// TIA Portal V20 program export: 0 tag tables, 36 data types, 10 data blocks, 80 code blocks (in call order from the OBs), 3 instance data blocks

TYPE "FRK_Access"
// stored: IsFailsafeCompliant false
   STRUCT
      CurrentLevel : DInt;
      CurrentUser : String[32];
      LoginFailed : Bool;
      Policy { S7_SetPoint := 'True'} : "ST_AccessPolicy";
      SessionGeneration : UDInt;
      LoginBusy : Bool;
      LoginResultSequence : UDInt;
      LoginTimeoutMs : UDInt;
      ProviderEnabled { ExternalAccessible := 'False'; ExternalVisible := 'False'; ExternalWritable := 'False'} : Bool;
      LastActivity { ExternalAccessible := 'False'; ExternalVisible := 'False'; ExternalWritable := 'False'} : UDInt;
      LoginSince { ExternalAccessible := 'False'; ExternalVisible := 'False'; ExternalWritable := 'False'} : UDInt;
      LoginSequence { ExternalAccessible := 'False'; ExternalVisible := 'False'; ExternalWritable := 'False'} : UDInt;
      CandidateUser { ExternalAccessible := 'False'; ExternalVisible := 'False'; ExternalWritable := 'False'} : String[32];
      CandidateLevel { ExternalAccessible := 'False'; ExternalVisible := 'False'; ExternalWritable := 'False'} : DInt;
      Round { ExternalAccessible := 'False'; ExternalVisible := 'False'; ExternalWritable := 'False'} : DInt;
      Salt { ExternalAccessible := 'False'; ExternalVisible := 'False'; ExternalWritable := 'False'} : Array[0..15] of Byte;
      Digest { ExternalAccessible := 'False'; ExternalVisible := 'False'; ExternalWritable := 'False'} : Array[0..31] of Byte;
      Expected { ExternalAccessible := 'False'; ExternalVisible := 'False'; ExternalWritable := 'False'} : Array[0..31] of Byte;
   END_STRUCT;
END_TYPE

TYPE "FRK_Carrier"
// stored: IsFailsafeCompliant false
   STRUCT
      Enabled { ExternalAccessible := 'False'; ExternalVisible := 'False'; ExternalWritable := 'False'} : Bool;
      Kind { ExternalAccessible := 'False'; ExternalVisible := 'False'; ExternalWritable := 'False'} : DInt;
      Serial { ExternalAccessible := 'False'; ExternalVisible := 'False'; ExternalWritable := 'False'} : UDInt;
      Context { ExternalAccessible := 'False'; ExternalVisible := 'False'; ExternalWritable := 'False'; S7_SetPoint := 'True'} : "ST_PartContext";
      Written { ExternalAccessible := 'False'; ExternalVisible := 'False'; ExternalWritable := 'False'; S7_SetPoint := 'True'} : "ST_PartContext";
      Writes { ExternalAccessible := 'False'; ExternalVisible := 'False'; ExternalWritable := 'False'} : UDInt;
   END_STRUCT;
END_TYPE

TYPE "FRK_ConfigCursor"
// stored: IsFailsafeCompliant false
   STRUCT
      Position { ExternalAccessible := 'False'; ExternalVisible := 'False'; ExternalWritable := 'False'} : DInt;
      First { ExternalAccessible := 'False'; ExternalVisible := 'False'; ExternalWritable := 'False'} : DInt;
   END_STRUCT;
END_TYPE

TYPE "FRK_Core"
// stored: IsFailsafeCompliant false
   STRUCT
      Named { ExternalAccessible := 'False'; ExternalVisible := 'False'; ExternalWritable := 'False'} : Bool;
      Initialized { ExternalAccessible := 'False'; ExternalVisible := 'False'; ExternalWritable := 'False'} : Bool;
      RegIndex { ExternalAccessible := 'False'; ExternalVisible := 'False'; ExternalWritable := 'False'} : DInt;
      ParentIndex { ExternalAccessible := 'False'; ExternalVisible := 'False'; ExternalWritable := 'False'} : DInt;
      ModuleType { ExternalAccessible := 'False'; ExternalVisible := 'False'; ExternalWritable := 'False'} : DInt;
      Exec { ExternalAccessible := 'False'; ExternalVisible := 'False'; ExternalWritable := 'False'} : DInt;
      ExecPrev { ExternalAccessible := 'False'; ExternalVisible := 'False'; ExternalWritable := 'False'} : Bool;
      AbortPrev { ExternalAccessible := 'False'; ExternalVisible := 'False'; ExternalWritable := 'False'} : Bool;
      Armed { ExternalAccessible := 'False'; ExternalVisible := 'False'; ExternalWritable := 'False'} : Bool;
      Command { ExternalAccessible := 'False'; ExternalVisible := 'False'; ExternalWritable := 'False'} : DInt;
      CommandLabel { ExternalAccessible := 'False'; ExternalVisible := 'False'; ExternalWritable := 'False'} : String[120];
      Dispatch { ExternalAccessible := 'False'; ExternalVisible := 'False'; ExternalWritable := 'False'} : Bool;
      EvInit { ExternalAccessible := 'False'; ExternalVisible := 'False'; ExternalWritable := 'False'} : Bool;
      EvCommandStart { ExternalAccessible := 'False'; ExternalVisible := 'False'; ExternalWritable := 'False'} : Bool;
      ReleasePending { ExternalAccessible := 'False'; ExternalVisible := 'False'; ExternalWritable := 'False'} : Bool;
      EvAbort { ExternalAccessible := 'False'; ExternalVisible := 'False'; ExternalWritable := 'False'} : Bool;
      EvAbortInError { ExternalAccessible := 'False'; ExternalVisible := 'False'; ExternalWritable := 'False'} : Bool;
      EvModeExit { ExternalAccessible := 'False'; ExternalVisible := 'False'; ExternalWritable := 'False'} : Bool;
      EvModeChanged { ExternalAccessible := 'False'; ExternalVisible := 'False'; ExternalWritable := 'False'} : Bool;
      "Step" { ExternalAccessible := 'False'; ExternalVisible := 'False'; ExternalWritable := 'False'} : DInt;
      HookResult { ExternalAccessible := 'False'; ExternalVisible := 'False'; ExternalWritable := 'False'} : DInt;
      Held { ExternalAccessible := 'False'; ExternalVisible := 'False'; ExternalWritable := 'False'} : Bool;
      HoldReq { ExternalAccessible := 'False'; ExternalVisible := 'False'; ExternalWritable := 'False'} : Bool;
      HoldReason { ExternalAccessible := 'False'; ExternalVisible := 'False'; ExternalWritable := 'False'} : DInt;
      DiagTouched { ExternalAccessible := 'False'; ExternalVisible := 'False'; ExternalWritable := 'False'} : Bool;
      TimingOpen { ExternalAccessible := 'False'; ExternalVisible := 'False'; ExternalWritable := 'False'} : Bool;
      StartMs { ExternalAccessible := 'False'; ExternalVisible := 'False'; ExternalWritable := 'False'} : UDInt;
      LastNowMs { ExternalAccessible := 'False'; ExternalVisible := 'False'; ExternalWritable := 'False'} : UDInt;
      DeltaMs { ExternalAccessible := 'False'; ExternalVisible := 'False'; ExternalWritable := 'False'} : UDInt;
      ActiveMs { ExternalAccessible := 'False'; ExternalVisible := 'False'; ExternalWritable := 'False'} : UDInt;
      TimeoutMs { ExternalAccessible := 'False'; ExternalVisible := 'False'; ExternalWritable := 'False'} : UDInt;
      Timing { ExternalAccessible := 'False'; ExternalVisible := 'False'; ExternalWritable := 'False'; S7_SetPoint := 'True'} : "ST_ModuleTiming";
   END_STRUCT;
END_TYPE

TYPE "FRK_ManualConditionRow"
// stored: IsFailsafeCompliant false
   STRUCT
      Used { ExternalAccessible := 'False'; ExternalVisible := 'False'; ExternalWritable := 'False'} : Bool;
      Value { ExternalAccessible := 'False'; ExternalVisible := 'False'; ExternalWritable := 'False'} : DInt;
      Ok { ExternalAccessible := 'False'; ExternalVisible := 'False'; ExternalWritable := 'False'} : Bool;
      Diag { ExternalAccessible := 'False'; ExternalVisible := 'False'; ExternalWritable := 'False'; S7_SetPoint := 'True'} : "ST_Diagnostic";
      Bypassable { ExternalAccessible := 'False'; ExternalVisible := 'False'; ExternalWritable := 'False'} : Bool;
   END_STRUCT;
END_TYPE

TYPE "FRK_RegistryRow"
// stored: IsFailsafeCompliant false
   STRUCT
      Valid { ExternalAccessible := 'False'; ExternalVisible := 'False'; ExternalWritable := 'False'} : Bool;
      Parent { ExternalAccessible := 'False'; ExternalVisible := 'False'; ExternalWritable := 'False'} : DInt;
      ModuleType { ExternalAccessible := 'False'; ExternalVisible := 'False'; ExternalWritable := 'False'} : DInt;
      TypeId { ExternalAccessible := 'False'; ExternalVisible := 'False'; ExternalWritable := 'False'} : DInt;
      Capabilities { ExternalAccessible := 'False'; ExternalVisible := 'False'; ExternalWritable := 'False'} : DWord;
      Exec { ExternalAccessible := 'False'; ExternalVisible := 'False'; ExternalWritable := 'False'} : DInt;
      ReasonCode { ExternalAccessible := 'False'; ExternalVisible := 'False'; ExternalWritable := 'False'} : DInt;
      Severity { ExternalAccessible := 'False'; ExternalVisible := 'False'; ExternalWritable := 'False'} : DInt;
   END_STRUCT;
END_TYPE

TYPE "FRK_Unit"
// stored: IsFailsafeCompliant false
   STRUCT
      Initialized { ExternalAccessible := 'False'; ExternalVisible := 'False'; ExternalWritable := 'False'} : Bool;
      Mode { ExternalAccessible := 'False'; ExternalVisible := 'False'; ExternalWritable := 'False'} : DInt;
      RequestedMode { ExternalAccessible := 'False'; ExternalVisible := 'False'; ExternalWritable := 'False'} : DInt;
      ModePending { ExternalAccessible := 'False'; ExternalVisible := 'False'; ExternalWritable := 'False'} : Bool;
      ExitFirst { ExternalAccessible := 'False'; ExternalVisible := 'False'; ExternalWritable := 'False'} : Bool;
      RunReq { ExternalAccessible := 'False'; ExternalVisible := 'False'; ExternalWritable := 'False'} : Bool;
      AbortReq { ExternalAccessible := 'False'; ExternalVisible := 'False'; ExternalWritable := 'False'} : Bool;
      StopReq { ExternalAccessible := 'False'; ExternalVisible := 'False'; ExternalWritable := 'False'} : Bool;
      ModeSince { ExternalAccessible := 'False'; ExternalVisible := 'False'; ExternalWritable := 'False'} : UDInt;
      ReleaseChildren { ExternalAccessible := 'False'; ExternalVisible := 'False'; ExternalWritable := 'False'} : Bool;
      Clearing { ExternalAccessible := 'False'; ExternalVisible := 'False'; ExternalWritable := 'False'} : Bool;
      FaultLatched { ExternalAccessible := 'False'; ExternalVisible := 'False'; ExternalWritable := 'False'} : Bool;
      PrevError { ExternalAccessible := 'False'; ExternalVisible := 'False'; ExternalWritable := 'False'} : Bool;
      EvReset { ExternalAccessible := 'False'; ExternalVisible := 'False'; ExternalWritable := 'False'} : Bool;
      SeenSequence { ExternalAccessible := 'False'; ExternalVisible := 'False'; ExternalWritable := 'False'} : UDInt;
      RequestPending { ExternalAccessible := 'False'; ExternalVisible := 'False'; ExternalWritable := 'False'} : Bool;
      Request { ExternalAccessible := 'False'; ExternalVisible := 'False'; ExternalWritable := 'False'; S7_SetPoint := 'True'} : "ST_HmiRequest";
      RequestUser { ExternalAccessible := 'False'; ExternalVisible := 'False'; ExternalWritable := 'False'} : String[32];
      Permit { ExternalAccessible := 'False'; ExternalVisible := 'False'; ExternalWritable := 'False'} : Bool;
      PermitDiag { ExternalAccessible := 'False'; ExternalVisible := 'False'; ExternalWritable := 'False'; S7_SetPoint := 'True'} : "ST_Diagnostic";
      CarrierIndex { ExternalAccessible := 'False'; ExternalVisible := 'False'; ExternalWritable := 'False'} : DInt;
      Good { ExternalAccessible := 'False'; ExternalVisible := 'False'; ExternalWritable := 'False'} : UDInt;
      Nok { ExternalAccessible := 'False'; ExternalVisible := 'False'; ExternalWritable := 'False'} : UDInt;
      Rework { ExternalAccessible := 'False'; ExternalVisible := 'False'; ExternalWritable := 'False'} : UDInt;
      NokReason { ExternalAccessible := 'False'; ExternalVisible := 'False'; ExternalWritable := 'False'} : DInt;
      CascadePending { ExternalAccessible := 'False'; ExternalVisible := 'False'; ExternalWritable := 'False'} : Bool;
      CascadeKind { ExternalAccessible := 'False'; ExternalVisible := 'False'; ExternalWritable := 'False'} : DInt;
      CascadeMode { ExternalAccessible := 'False'; ExternalVisible := 'False'; ExternalWritable := 'False'} : DInt;
      FollowStart { ExternalAccessible := 'False'; ExternalVisible := 'False'; ExternalWritable := 'False'} : Bool;
   END_STRUCT;
END_TYPE

TYPE "ST_AccessPolicy"
// stored: IsFailsafeCompliant false
   STRUCT
      Required : Array[0..11] of DInt;
      SessionTimeout : Time := T#0MS;
   END_STRUCT;
END_TYPE

TYPE "ST_CommandInfo"
// stored: IsFailsafeCompliant false
   STRUCT
      Value : DInt;
      Label : String[120];
      Style : DInt;
   END_STRUCT;
END_TYPE

TYPE "ST_ConfigEntry"
// stored: IsFailsafeCompliant false
   STRUCT
      Scope : WString[255];
      Item : WString[255];
      ValueText : WString[255];
      WriteKey : String[160];
      WriteRevision : UDInt;
      ConfigKind : DInt;
      ValueType : DInt;
      Writable : Bool;
      RequiresReady : Bool;
      HasMinimum : Bool;
      HasMaximum : Bool;
      Minimum : LReal;
      Maximum : LReal;
      Unit : String[16];
      LabelKey : String[160];
      EnumDomain : WString[255];
      ClassId : String[40];
      ReadLevel : DInt;
      WriteLevel : DInt;
      Readable : Bool;
      UnitCode : DInt;
      EnumLabelKey : String[80];
      ModelScoped : Bool;
   END_STRUCT;
END_TYPE

TYPE "ST_ConfigPage"
// stored: IsFailsafeCompliant false
   STRUCT
      Revision : UDInt;
      PageIndex : Int;
      PageCount : Int;
      EntryCount : Int;
      Entries { S7_SetPoint := 'True'} : Array[1..16] of "ST_ConfigEntry";
   END_STRUCT;
END_TYPE

TYPE "ST_DeclarationCellHal"
// stored: IsFailsafeCompliant false
   STRUCT
      Clamp { ExternalAccessible := 'False'; ExternalVisible := 'False'; ExternalWritable := 'False'; S7_SetPoint := 'True'} : "ST_DeclarationLeafHal";
      Gate { ExternalAccessible := 'False'; ExternalVisible := 'False'; ExternalWritable := 'False'; S7_SetPoint := 'True'} : "ST_DeclarationLeafHal";
   END_STRUCT;
END_TYPE

TYPE "ST_DeclarationLeafHal"
// stored: IsFailsafeCompliant false
   STRUCT
      Sample : DInt;
      Permit : Bool := TRUE;
      Finish : Bool;
      BackgroundFault : Bool;
      Diag { S7_SetPoint := 'True'} : "ST_Diagnostic";
      LaterDiag { S7_SetPoint := 'True'} : "ST_Diagnostic";
      ExitHold : Bool;
      Verdict : DInt := 1;
   END_STRUCT;
END_TYPE

TYPE "ST_DeclarationOutCmd"
// stored: IsFailsafeCompliant false
   STRUCT
      Result : DInt;
   END_STRUCT;
END_TYPE

TYPE "ST_DeclarationOutImm"
// stored: IsFailsafeCompliant false
   STRUCT
      Sample : DInt;
      InitCount : DInt;
      StartCount : DInt;
      CyclicCount : DInt;
      AbortCount : DInt;
      ErrorAbortCount : DInt;
      DispatchCount : DInt;
      SeenValue : DInt;
      Ordered : Bool;
      Output : Bool;
   END_STRUCT;
END_TYPE

TYPE "ST_DeclarationParCfg"
// stored: IsFailsafeCompliant false
   STRUCT
      SchemaVersion : UInt := 3;
      Timeout : Time := T#2S;
   END_STRUCT;
END_TYPE

TYPE "ST_DeclarationParCmd"
// stored: IsFailsafeCompliant false
   STRUCT
      Value : DInt;
   END_STRUCT;
END_TYPE

TYPE "ST_DeclarationUnitHal"
// stored: IsFailsafeCompliant false
   STRUCT
      Cell { ExternalAccessible := 'False'; ExternalVisible := 'False'; ExternalWritable := 'False'; S7_SetPoint := 'True'} : "ST_DeclarationCellHal";
      Satellite { ExternalAccessible := 'False'; ExternalVisible := 'False'; ExternalWritable := 'False'; S7_SetPoint := 'True'} : "ST_SatelliteUnitHal";
   END_STRUCT;
END_TYPE

TYPE "ST_Diagnostic"
// stored: IsFailsafeCompliant false
   STRUCT
      ReasonCode : DInt;
      SourcePath : WString[255];
      Description : WString[255];
      IoTag : String[80];
      IoAddress : String[80];
      Severity : DInt;
      Category : DInt;
      Since : LDT;
      TimeSynchronized : Bool;
   END_STRUCT;
END_TYPE

TYPE "ST_FraktalHal"
// stored: IsFailsafeCompliant false
   STRUCT
      StationA { ExternalAccessible := 'False'; ExternalVisible := 'False'; ExternalWritable := 'False'; S7_SetPoint := 'True'} : "ST_DeclarationUnitHal";
      StationB { ExternalAccessible := 'False'; ExternalVisible := 'False'; ExternalWritable := 'False'; S7_SetPoint := 'True'} : "ST_DeclarationUnitHal";
   END_STRUCT;
END_TYPE

TYPE "ST_HmiRequest"
// stored: IsFailsafeCompliant false
   STRUCT
      Kind : DInt;
      TargetPath : WString[255];
      NameValue : String[160];
      TextValue : WString[255];
      User : String[32];
      Secret : String[32];
      IntValue : DInt;
      BoolValue : Bool;
      DurationMs : UDInt;
      Sequence : UDInt;
   END_STRUCT;
END_TYPE

TYPE "ST_HmiResponse"
// stored: IsFailsafeCompliant false
   STRUCT
      AckSequence : UDInt;
      Accepted : Bool;
      Diagnostic : WString[255];
      Report { S7_SetPoint := 'True'} : "ST_ReleaseReport";
      ConfigPage { S7_SetPoint := 'True'} : "ST_ConfigPage";
   END_STRUCT;
END_TYPE

TYPE "ST_InnerUnitHal"
// stored: IsFailsafeCompliant false
   STRUCT
      Cell { ExternalAccessible := 'False'; ExternalVisible := 'False'; ExternalWritable := 'False'; S7_SetPoint := 'True'} : "ST_DeclarationCellHal";
   END_STRUCT;
END_TYPE

TYPE "ST_MeasRecord"
// stored: IsFailsafeCompliant false
   STRUCT
      "Name" : String[64];
      Value : LReal;
      Minimum : LReal;
      Maximum : LReal;
      Target : LReal;
      Unit : String[16];
      InTol : Bool;
   END_STRUCT;
END_TYPE

TYPE "ST_ModePolicy"
// stored: IsFailsafeCompliant false
   STRUCT
      Shield : DInt;
      Style : DInt;
   END_STRUCT;
END_TYPE

TYPE "ST_ModuleStatus"
// stored: IsFailsafeCompliant false
   STRUCT
      "Name" : String[80];
      DisplayNameKey : String[160];
      DescriptionKey : String[160];
      TypeKey : String[160];
      ModuleType : DInt;
      State : DInt;
      FaultActive : Bool;
      Diagnostic { S7_SetPoint := 'True'} : "ST_Diagnostic";
      TileEnable : Bool := TRUE;
      ControlDomainId : String[80];
   END_STRUCT;
END_TYPE

TYPE "ST_ModuleTiming"
// stored: IsFailsafeCompliant false
   STRUCT
      LastCmdTime : Time;
      Rows { S7_SetPoint := 'True'} : Array[1..8] of "ST_TimingRow";
      Truncated : Bool;
   END_STRUCT;
END_TYPE

TYPE "ST_PartContext"
// stored: IsFailsafeCompliant false
   STRUCT
      Uid : String[64];
      Present : Bool;
      CarrierKind : DInt;
      Result { S7_SetPoint := 'True'} : "ST_PartResult";
      Parents : Array[1..8] of String[64];
   END_STRUCT;
END_TYPE

TYPE "ST_PartResult"
// stored: IsFailsafeCompliant false
   STRUCT
      Verdict : DInt;
      ReasonCode : DInt;
      Records { S7_SetPoint := 'True'} : Array[1..32] of "ST_MeasRecord";
      StationPath : WString[255];
      Stamp : LDT;
      TimeSynchronized : Bool;
   END_STRUCT;
END_TYPE

TYPE "ST_ReleaseReason"
// stored: IsFailsafeCompliant false
   STRUCT
      Description : WString[255];
      ReasonCode : DInt;
      SourcePath : WString[255];
      Kind : DInt;
      Bypassable : Bool;
   END_STRUCT;
END_TYPE

TYPE "ST_ReleaseReport"
// stored: IsFailsafeCompliant false
   STRUCT
      Released : Bool;
      Count : Int;
      Reasons { S7_SetPoint := 'True'} : Array[1..24] of "ST_ReleaseReason";
   END_STRUCT;
END_TYPE

TYPE "ST_SatelliteUnitHal"
// stored: IsFailsafeCompliant false
   STRUCT
      Cell { ExternalAccessible := 'False'; ExternalVisible := 'False'; ExternalWritable := 'False'; S7_SetPoint := 'True'} : "ST_DeclarationCellHal";
      Inner { ExternalAccessible := 'False'; ExternalVisible := 'False'; ExternalWritable := 'False'; S7_SetPoint := 'True'} : "ST_InnerUnitHal";
   END_STRUCT;
END_TYPE

TYPE "ST_TimingRow"
// stored: IsFailsafeCompliant false
   STRUCT
      Id : DInt;
      Label : String[120];
      TimeClass : DInt;
      Count : UDInt;
      Last : Time;
      Minimum : Time;
      Maximum : Time;
      Avg : Time;
   END_STRUCT;
END_TYPE

TYPE "ST_UnitProbeDevice"
// stored: IsFailsafeCompliant false
   STRUCT
      Cycles : UDInt;
      ExitCalls : UDInt;
      Changes : UDInt;
      Resets : UDInt;
      Received : Bool;
      Processed : Bool;
   END_STRUCT;
END_TYPE

TYPE "ST_UnitProbeImm"
// stored: IsFailsafeCompliant false
   STRUCT
      Cycles : UDInt;
      ExitCalls : UDInt;
      Changes : UDInt;
      Resets : UDInt;
   END_STRUCT;
END_TYPE

TYPE "ST_UserRecord"
// stored: IsFailsafeCompliant false
   STRUCT
      User : String[32];
      Salt : Array[0..15] of Byte;
      PinHash : Array[0..31] of Byte;
      Level : DInt;
   END_STRUCT;
END_TYPE

DATA_BLOCK "FRK_Carriers"   // DB3
{ S7_Optimized_Access := 'TRUE' }
VERSION : 0.1
// stored: AutoNumber true, DBAccessibleFromOPCUA true, DBAccessibleFromWebserver true, IsOnlyStoredInLoadMemory false, IsRetainMemResEnabled false, IsWriteProtectedInAS false, MemoryReserve 100
   VAR
      Slots { ExternalAccessible := 'False'; ExternalVisible := 'False'; ExternalWritable := 'False'; S7_SetPoint := 'True'} : Array[0..32] of "FRK_Carrier";
   END_VAR
BEGIN
END_DATA_BLOCK

DATA_BLOCK "FRK_Clock"   // DB1
{ S7_Optimized_Access := 'TRUE' }
VERSION : 0.1
// stored: AutoNumber true, DBAccessibleFromOPCUA true, DBAccessibleFromWebserver true, IsOnlyStoredInLoadMemory false, IsRetainMemResEnabled false, IsWriteProtectedInAS false, MemoryReserve 100
   VAR
      Mem { ExternalAccessible := 'False'; ExternalVisible := 'False'; ExternalWritable := 'False'} : LReal;
      AccMs { ExternalAccessible := 'False'; ExternalVisible := 'False'; ExternalWritable := 'False'} : LReal;
      NowMs { ExternalAccessible := 'False'; ExternalVisible := 'False'; ExternalWritable := 'False'} : UDInt;
   END_VAR
BEGIN
END_DATA_BLOCK

DATA_BLOCK "FRK_LocalUsers"   // DB4
{ S7_Optimized_Access := 'TRUE' }
VERSION : 0.1
// stored: AutoNumber true, DBAccessibleFromOPCUA true, DBAccessibleFromWebserver true, IsOnlyStoredInLoadMemory false, IsRetainMemResEnabled false, IsWriteProtectedInAS false, MemoryReserve 100
   VAR
      Count { ExternalAccessible := 'False'; ExternalVisible := 'False'; ExternalWritable := 'False'} : DInt;
      Rows { ExternalAccessible := 'False'; ExternalVisible := 'False'; ExternalWritable := 'False'; S7_SetPoint := 'True'} : Array[1..16] of "ST_UserRecord";
   END_VAR
BEGIN
END_DATA_BLOCK

DATA_BLOCK "FRK_Registry"   // DB2
{ S7_Optimized_Access := 'TRUE' }
VERSION : 0.1
// stored: AutoNumber true, DBAccessibleFromOPCUA true, DBAccessibleFromWebserver true, IsOnlyStoredInLoadMemory false, IsRetainMemResEnabled false, IsWriteProtectedInAS false, MemoryReserve 100
   VAR
      Count { ExternalAccessible := 'False'; ExternalVisible := 'False'; ExternalWritable := 'False'} : DInt;
      Fault { ExternalAccessible := 'False'; ExternalVisible := 'False'; ExternalWritable := 'False'} : Bool;
      Rows { ExternalAccessible := 'False'; ExternalVisible := 'False'; ExternalWritable := 'False'; S7_SetPoint := 'True'} : Array[0..32] of "FRK_RegistryRow";
   END_VAR
BEGIN
END_DATA_BLOCK

DATA_BLOCK "FRK_UnitScratch"   // DB5
{ S7_Optimized_Access := 'TRUE' }
VERSION : 0.1
// stored: AutoNumber true, DBAccessibleFromOPCUA true, DBAccessibleFromWebserver true, IsOnlyStoredInLoadMemory false, IsRetainMemResEnabled false, IsWriteProtectedInAS false, MemoryReserve 100
   VAR
      Response { ExternalAccessible := 'False'; ExternalVisible := 'False'; ExternalWritable := 'False'; S7_SetPoint := 'True'} : "ST_HmiResponse";
      EmptyDiagnostic { ExternalAccessible := 'False'; ExternalVisible := 'False'; ExternalWritable := 'False'; S7_SetPoint := 'True'} : "ST_Diagnostic";
      EmptyConfigEntry { ExternalAccessible := 'False'; ExternalVisible := 'False'; ExternalWritable := 'False'; S7_SetPoint := 'True'} : "ST_ConfigEntry";
   END_VAR
BEGIN
END_DATA_BLOCK

DATA_BLOCK "GDB_AccessTest"   // DB6
{ S7_Optimized_Access := 'TRUE' }
VERSION : 0.1
// stored: AutoNumber true, DBAccessibleFromOPCUA true, DBAccessibleFromWebserver true, IsOnlyStoredInLoadMemory false, IsRetainMemResEnabled false, IsWriteProtectedInAS false, MemoryReserve 100
   VAR
      ProviderOff : Bool;
      CancelOnLogin : Bool;
      SupersedeOnLogin : Bool;
      InterruptedBusy { ExternalWritable := 'False'} : Bool;
      SupersededSequence { ExternalWritable := 'False'} : UDInt;
      InterruptRequest { ExternalAccessible := 'False'; ExternalVisible := 'False'; ExternalWritable := 'False'; S7_SetPoint := 'True'} : "ST_HmiRequest";
      HashData { ExternalAccessible := 'False'; ExternalVisible := 'False'; ExternalWritable := 'False'} : Array[0..47] of Byte;
      Hash0 { ExternalWritable := 'False'} : Array[0..31] of Byte;
      Hash1 { ExternalWritable := 'False'} : Array[0..31] of Byte;
      Hash2 { ExternalWritable := 'False'} : Array[0..31] of Byte;
      Hash3 { ExternalWritable := 'False'} : Array[0..31] of Byte;
      HashOk { ExternalWritable := 'False'} : Bool;
   END_VAR
BEGIN
END_DATA_BLOCK

DATA_BLOCK "GDB_FraktalHal"   // DB10
{ S7_Optimized_Access := 'TRUE' }
VERSION : 0.1
// stored: AutoNumber true, DBAccessibleFromOPCUA true, DBAccessibleFromWebserver true, IsOnlyStoredInLoadMemory false, IsRetainMemResEnabled false, IsWriteProtectedInAS false, MemoryReserve 100
   VAR
      Data { ExternalAccessible := 'False'; ExternalVisible := 'False'; ExternalWritable := 'False'; S7_SetPoint := 'True'} : "ST_FraktalHal";
   END_VAR
BEGIN
END_DATA_BLOCK

DATA_BLOCK "GDB_ManifestTest"   // DB7
{ S7_Optimized_Access := 'TRUE' }
VERSION : 0.1
// stored: AutoNumber true, DBAccessibleFromOPCUA true, DBAccessibleFromWebserver true, IsOnlyStoredInLoadMemory false, IsRetainMemResEnabled false, IsWriteProtectedInAS false, MemoryReserve 100
   VAR
      ReadLock : Bool;
   END_VAR
BEGIN
END_DATA_BLOCK

DATA_BLOCK "GDB_RoutingTest"   // DB8
{ S7_Optimized_Access := 'TRUE' }
VERSION : 0.1
// stored: AutoNumber true, DBAccessibleFromOPCUA true, DBAccessibleFromWebserver true, IsOnlyStoredInLoadMemory false, IsRetainMemResEnabled false, IsWriteProtectedInAS false, MemoryReserve 100
   VAR
      PermitOne : Bool;
      PermitTwo : Bool;
      NestedFinish : Bool;
      InnerFinish : Bool;
      NestedAccessLock : Bool;
      RootManualPermit : Bool;
      ManualAccessLock : Bool;
      LocalPulse : Bool;
      LocalKind : DInt;
      LocalValue : DInt;
      LocalAccepted { ExternalWritable := 'False'} : Bool;
      LocalFirstKind { ExternalWritable := 'False'} : DInt;
      LocalRequest { ExternalAccessible := 'False'; ExternalVisible := 'False'; ExternalWritable := 'False'; S7_SetPoint := 'True'} : "ST_HmiRequest";
      ManExecute { ExternalWritable := 'False'} : Bool;
      ManStarts { ExternalWritable := 'False'} : DInt;
   END_VAR
BEGIN
END_DATA_BLOCK

DATA_BLOCK "GDB_UnitTest"   // DB9
{ S7_Optimized_Access := 'TRUE' }
VERSION : 0.1
// stored: AutoNumber true, DBAccessibleFromOPCUA true, DBAccessibleFromWebserver true, IsOnlyStoredInLoadMemory false, IsRetainMemResEnabled false, IsWriteProtectedInAS false, MemoryReserve 100
   VAR
      FinishCycle : Bool;
      Permit : Bool;
      FaultRoot : Bool;
      ExitHold : Bool;
      LockStart : Bool;
      IssueChild : Bool;
      ChildCommand : DInt;
      Verdict : DInt;
      Reason : DInt;
      CarrierControl : DInt;
      Scans { ExternalWritable := 'False'} : UDInt;
      Restarts { ExternalWritable := 'False'} : UDInt;
      ChildExecute { ExternalWritable := 'False'} : Bool;
      ChildState { ExternalWritable := 'False'} : DInt;
      CarrierWrites { ExternalWritable := 'False'} : UDInt;
      CarrierSerial { ExternalWritable := 'False'} : UDInt;
      WrittenUid { ExternalWritable := 'False'} : String[64];
      WrittenVerdict { ExternalWritable := 'False'} : DInt;
      LastEvent { ExternalWritable := 'False'} : DInt;
      SecretCleared { ExternalWritable := 'False'} : Bool;
      SnapshotSecretCleared { ExternalWritable := 'False'} : Bool;
      BootStamp { ExternalWritable := 'False'} : LDT;
   END_VAR
BEGIN
END_DATA_BLOCK

ORGANIZATION_BLOCK "Main"   // OB1, SCL, ProgramCycle
{ S7_Optimized_Access := 'TRUE' }
VERSION : 0.1
// stored: AutoNumber true, IsIECCheckEnabled false, SetENOAutomatically false
   VAR_INPUT
      Initial_Call : Bool;   // Initial call of this OB
      Remanence : Bool;   // =True, if remanent data are available
   END_VAR
   VAR_TEMP
      StartupStamp : DTL;
      ResultCode : Int;
   END_VAR
BEGIN

   IF #Initial_Call THEN
       "FRK_LocalUsers".Count := 2;
       "FRK_LocalUsers".Rows[1].User := 'operator';
       "FRK_LocalUsers".Rows[1].Level := 1;
       "FRK_LocalUsers".Rows[1].Salt[0] := BYTE#16#10;
       "FRK_LocalUsers".Rows[1].Salt[1] := BYTE#16#BD;
       "FRK_LocalUsers".Rows[1].Salt[2] := BYTE#16#42;
       "FRK_LocalUsers".Rows[1].Salt[3] := BYTE#16#1E;
       "FRK_LocalUsers".Rows[1].Salt[4] := BYTE#16#34;
       "FRK_LocalUsers".Rows[1].Salt[5] := BYTE#16#C3;
       "FRK_LocalUsers".Rows[1].Salt[6] := BYTE#16#71;
       "FRK_LocalUsers".Rows[1].Salt[7] := BYTE#16#89;
       "FRK_LocalUsers".Rows[1].Salt[8] := BYTE#16#CF;
       "FRK_LocalUsers".Rows[1].Salt[9] := BYTE#16#68;
       "FRK_LocalUsers".Rows[1].Salt[10] := BYTE#16#93;
       "FRK_LocalUsers".Rows[1].Salt[11] := BYTE#16#47;
       "FRK_LocalUsers".Rows[1].Salt[12] := BYTE#16#BB;
       "FRK_LocalUsers".Rows[1].Salt[13] := BYTE#16#CB;
       "FRK_LocalUsers".Rows[1].Salt[14] := BYTE#16#DB;
       "FRK_LocalUsers".Rows[1].Salt[15] := BYTE#16#1B;
       "FRK_LocalUsers".Rows[1].PinHash[0] := BYTE#16#EB;
       "FRK_LocalUsers".Rows[1].PinHash[1] := BYTE#16#77;
       "FRK_LocalUsers".Rows[1].PinHash[2] := BYTE#16#28;
       "FRK_LocalUsers".Rows[1].PinHash[3] := BYTE#16#BE;
       "FRK_LocalUsers".Rows[1].PinHash[4] := BYTE#16#AA;
       "FRK_LocalUsers".Rows[1].PinHash[5] := BYTE#16#21;
       "FRK_LocalUsers".Rows[1].PinHash[6] := BYTE#16#75;
       "FRK_LocalUsers".Rows[1].PinHash[7] := BYTE#16#34;
       "FRK_LocalUsers".Rows[1].PinHash[8] := BYTE#16#91;
       "FRK_LocalUsers".Rows[1].PinHash[9] := BYTE#16#8C;
       "FRK_LocalUsers".Rows[1].PinHash[10] := BYTE#16#F2;
       "FRK_LocalUsers".Rows[1].PinHash[11] := BYTE#16#B5;
       "FRK_LocalUsers".Rows[1].PinHash[12] := BYTE#16#63;
       "FRK_LocalUsers".Rows[1].PinHash[13] := BYTE#16#85;
       "FRK_LocalUsers".Rows[1].PinHash[14] := BYTE#16#28;
       "FRK_LocalUsers".Rows[1].PinHash[15] := BYTE#16#DF;
       "FRK_LocalUsers".Rows[1].PinHash[16] := BYTE#16#0D;
       "FRK_LocalUsers".Rows[1].PinHash[17] := BYTE#16#AA;
       "FRK_LocalUsers".Rows[1].PinHash[18] := BYTE#16#59;
       "FRK_LocalUsers".Rows[1].PinHash[19] := BYTE#16#4E;
       "FRK_LocalUsers".Rows[1].PinHash[20] := BYTE#16#93;
       "FRK_LocalUsers".Rows[1].PinHash[21] := BYTE#16#6B;
       "FRK_LocalUsers".Rows[1].PinHash[22] := BYTE#16#43;
       "FRK_LocalUsers".Rows[1].PinHash[23] := BYTE#16#85;
       "FRK_LocalUsers".Rows[1].PinHash[24] := BYTE#16#7F;
       "FRK_LocalUsers".Rows[1].PinHash[25] := BYTE#16#1F;
       "FRK_LocalUsers".Rows[1].PinHash[26] := BYTE#16#D4;
       "FRK_LocalUsers".Rows[1].PinHash[27] := BYTE#16#7C;
       "FRK_LocalUsers".Rows[1].PinHash[28] := BYTE#16#68;
       "FRK_LocalUsers".Rows[1].PinHash[29] := BYTE#16#26;
       "FRK_LocalUsers".Rows[1].PinHash[30] := BYTE#16#EE;
       "FRK_LocalUsers".Rows[1].PinHash[31] := BYTE#16#68;
       "FRK_LocalUsers".Rows[2].User := 'admin';
       "FRK_LocalUsers".Rows[2].Level := 4;
       "FRK_LocalUsers".Rows[2].Salt[0] := BYTE#16#86;
       "FRK_LocalUsers".Rows[2].Salt[1] := BYTE#16#55;
       "FRK_LocalUsers".Rows[2].Salt[2] := BYTE#16#D5;
       "FRK_LocalUsers".Rows[2].Salt[3] := BYTE#16#84;
       "FRK_LocalUsers".Rows[2].Salt[4] := BYTE#16#27;
       "FRK_LocalUsers".Rows[2].Salt[5] := BYTE#16#D6;
       "FRK_LocalUsers".Rows[2].Salt[6] := BYTE#16#72;
       "FRK_LocalUsers".Rows[2].Salt[7] := BYTE#16#35;
       "FRK_LocalUsers".Rows[2].Salt[8] := BYTE#16#F8;
       "FRK_LocalUsers".Rows[2].Salt[9] := BYTE#16#F1;
       "FRK_LocalUsers".Rows[2].Salt[10] := BYTE#16#A3;
       "FRK_LocalUsers".Rows[2].Salt[11] := BYTE#16#B6;
       "FRK_LocalUsers".Rows[2].Salt[12] := BYTE#16#EC;
       "FRK_LocalUsers".Rows[2].Salt[13] := BYTE#16#77;
       "FRK_LocalUsers".Rows[2].Salt[14] := BYTE#16#E2;
       "FRK_LocalUsers".Rows[2].Salt[15] := BYTE#16#CB;
       "FRK_LocalUsers".Rows[2].PinHash[0] := BYTE#16#CB;
       "FRK_LocalUsers".Rows[2].PinHash[1] := BYTE#16#99;
       "FRK_LocalUsers".Rows[2].PinHash[2] := BYTE#16#67;
       "FRK_LocalUsers".Rows[2].PinHash[3] := BYTE#16#9C;
       "FRK_LocalUsers".Rows[2].PinHash[4] := BYTE#16#33;
       "FRK_LocalUsers".Rows[2].PinHash[5] := BYTE#16#4D;
       "FRK_LocalUsers".Rows[2].PinHash[6] := BYTE#16#6C;
       "FRK_LocalUsers".Rows[2].PinHash[7] := BYTE#16#50;
       "FRK_LocalUsers".Rows[2].PinHash[8] := BYTE#16#EE;
       "FRK_LocalUsers".Rows[2].PinHash[9] := BYTE#16#AB;
       "FRK_LocalUsers".Rows[2].PinHash[10] := BYTE#16#B2;
       "FRK_LocalUsers".Rows[2].PinHash[11] := BYTE#16#26;
       "FRK_LocalUsers".Rows[2].PinHash[12] := BYTE#16#A8;
       "FRK_LocalUsers".Rows[2].PinHash[13] := BYTE#16#7A;
       "FRK_LocalUsers".Rows[2].PinHash[14] := BYTE#16#07;
       "FRK_LocalUsers".Rows[2].PinHash[15] := BYTE#16#0A;
       "FRK_LocalUsers".Rows[2].PinHash[16] := BYTE#16#3D;
       "FRK_LocalUsers".Rows[2].PinHash[17] := BYTE#16#8A;
       "FRK_LocalUsers".Rows[2].PinHash[18] := BYTE#16#03;
       "FRK_LocalUsers".Rows[2].PinHash[19] := BYTE#16#9E;
       "FRK_LocalUsers".Rows[2].PinHash[20] := BYTE#16#9C;
       "FRK_LocalUsers".Rows[2].PinHash[21] := BYTE#16#EA;
       "FRK_LocalUsers".Rows[2].PinHash[22] := BYTE#16#A3;
       "FRK_LocalUsers".Rows[2].PinHash[23] := BYTE#16#47;
       "FRK_LocalUsers".Rows[2].PinHash[24] := BYTE#16#DE;
       "FRK_LocalUsers".Rows[2].PinHash[25] := BYTE#16#0B;
       "FRK_LocalUsers".Rows[2].PinHash[26] := BYTE#16#B7;
       "FRK_LocalUsers".Rows[2].PinHash[27] := BYTE#16#38;
       "FRK_LocalUsers".Rows[2].PinHash[28] := BYTE#16#0F;
       "FRK_LocalUsers".Rows[2].PinHash[29] := BYTE#16#22;
       "FRK_LocalUsers".Rows[2].PinHash[30] := BYTE#16#F0;
       "FRK_LocalUsers".Rows[2].PinHash[31] := BYTE#16#D4;
       "StationA".Access.Policy.Required[2] := 1;
       "StationA".Access.Policy.Required[4] := 1;
       "StationA".Access.Policy.Required[5] := 1;
       "StationA".Access.Policy.Required[8] := 4;
       "StationA".Access.Policy.SessionTimeout := T#0ms;
       "StationB".Access.Policy.Required[2] := 1;
       "StationB".Access.Policy.Required[4] := 1;
       "StationB".Access.Policy.Required[5] := 1;
       "StationB".Access.Policy.Required[8] := 4;
       "StationB".Access.Policy.SessionTimeout := T#0ms;
       "GDB_AccessTest".HashData[0] := BYTE#16#00;
       "GDB_AccessTest".HashData[1] := BYTE#16#01;
       "GDB_AccessTest".HashData[2] := BYTE#16#02;
       "GDB_AccessTest".HashData[3] := BYTE#16#03;
       "GDB_AccessTest".HashData[4] := BYTE#16#04;
       "GDB_AccessTest".HashData[5] := BYTE#16#05;
       "GDB_AccessTest".HashData[6] := BYTE#16#06;
       "GDB_AccessTest".HashData[7] := BYTE#16#07;
       "GDB_AccessTest".HashData[8] := BYTE#16#08;
       "GDB_AccessTest".HashData[9] := BYTE#16#09;
       "GDB_AccessTest".HashData[10] := BYTE#16#0A;
       "GDB_AccessTest".HashData[11] := BYTE#16#0B;
       "GDB_AccessTest".HashData[12] := BYTE#16#0C;
       "GDB_AccessTest".HashData[13] := BYTE#16#0D;
       "GDB_AccessTest".HashData[14] := BYTE#16#0E;
       "GDB_AccessTest".HashData[15] := BYTE#16#0F;
       "GDB_AccessTest".HashData[16] := BYTE#16#10;
       "GDB_AccessTest".HashData[17] := BYTE#16#11;
       "GDB_AccessTest".HashData[18] := BYTE#16#12;
       "GDB_AccessTest".HashData[19] := BYTE#16#13;
       "GDB_AccessTest".HashData[20] := BYTE#16#14;
       "GDB_AccessTest".HashData[21] := BYTE#16#15;
       "GDB_AccessTest".HashData[22] := BYTE#16#16;
       "GDB_AccessTest".HashData[23] := BYTE#16#17;
       "GDB_AccessTest".HashData[24] := BYTE#16#18;
       "GDB_AccessTest".HashData[25] := BYTE#16#19;
       "GDB_AccessTest".HashData[26] := BYTE#16#1A;
       "GDB_AccessTest".HashData[27] := BYTE#16#1B;
       "GDB_AccessTest".HashData[28] := BYTE#16#1C;
       "GDB_AccessTest".HashData[29] := BYTE#16#1D;
       "GDB_AccessTest".HashData[30] := BYTE#16#1E;
       "GDB_AccessTest".HashData[31] := BYTE#16#1F;
       "GDB_AccessTest".HashData[32] := BYTE#16#20;
       "GDB_AccessTest".HashData[33] := BYTE#16#21;
       "GDB_AccessTest".HashData[34] := BYTE#16#22;
       "GDB_AccessTest".HashData[35] := BYTE#16#23;
       "GDB_AccessTest".HashData[36] := BYTE#16#24;
       "GDB_AccessTest".HashData[37] := BYTE#16#25;
       "GDB_AccessTest".HashData[38] := BYTE#16#26;
       "GDB_AccessTest".HashData[39] := BYTE#16#27;
       "GDB_AccessTest".HashData[40] := BYTE#16#28;
       "GDB_AccessTest".HashData[41] := BYTE#16#29;
       "GDB_AccessTest".HashData[42] := BYTE#16#2A;
       "GDB_AccessTest".HashData[43] := BYTE#16#2B;
       "GDB_AccessTest".HashData[44] := BYTE#16#2C;
       "GDB_AccessTest".HashData[45] := BYTE#16#2D;
       "GDB_AccessTest".HashData[46] := BYTE#16#2E;
       "GDB_AccessTest".HashData[47] := BYTE#16#2F;
       "GDB_AccessTest".HashOk := "FRK_Sha256Pin"(Data := "GDB_AccessTest".HashData, Size := 0, Digest := "GDB_AccessTest".Hash0);
       "GDB_AccessTest".HashData[0] := BYTE#16#61;
       "GDB_AccessTest".HashData[1] := BYTE#16#62;
       "GDB_AccessTest".HashData[2] := BYTE#16#63;
       "GDB_AccessTest".HashData[3] := BYTE#16#00;
       "GDB_AccessTest".HashData[4] := BYTE#16#00;
       "GDB_AccessTest".HashData[5] := BYTE#16#00;
       "GDB_AccessTest".HashData[6] := BYTE#16#00;
       "GDB_AccessTest".HashData[7] := BYTE#16#00;
       "GDB_AccessTest".HashData[8] := BYTE#16#00;
       "GDB_AccessTest".HashData[9] := BYTE#16#00;
       "GDB_AccessTest".HashData[10] := BYTE#16#00;
       "GDB_AccessTest".HashData[11] := BYTE#16#00;
       "GDB_AccessTest".HashData[12] := BYTE#16#00;
       "GDB_AccessTest".HashData[13] := BYTE#16#00;
       "GDB_AccessTest".HashData[14] := BYTE#16#00;
       "GDB_AccessTest".HashData[15] := BYTE#16#00;
       "GDB_AccessTest".HashData[16] := BYTE#16#00;
       "GDB_AccessTest".HashData[17] := BYTE#16#00;
       "GDB_AccessTest".HashData[18] := BYTE#16#00;
       "GDB_AccessTest".HashData[19] := BYTE#16#00;
       "GDB_AccessTest".HashData[20] := BYTE#16#00;
       "GDB_AccessTest".HashData[21] := BYTE#16#00;
       "GDB_AccessTest".HashData[22] := BYTE#16#00;
       "GDB_AccessTest".HashData[23] := BYTE#16#00;
       "GDB_AccessTest".HashData[24] := BYTE#16#00;
       "GDB_AccessTest".HashData[25] := BYTE#16#00;
       "GDB_AccessTest".HashData[26] := BYTE#16#00;
       "GDB_AccessTest".HashData[27] := BYTE#16#00;
       "GDB_AccessTest".HashData[28] := BYTE#16#00;
       "GDB_AccessTest".HashData[29] := BYTE#16#00;
       "GDB_AccessTest".HashData[30] := BYTE#16#00;
       "GDB_AccessTest".HashData[31] := BYTE#16#00;
       "GDB_AccessTest".HashData[32] := BYTE#16#00;
       "GDB_AccessTest".HashData[33] := BYTE#16#00;
       "GDB_AccessTest".HashData[34] := BYTE#16#00;
       "GDB_AccessTest".HashData[35] := BYTE#16#00;
       "GDB_AccessTest".HashData[36] := BYTE#16#00;
       "GDB_AccessTest".HashData[37] := BYTE#16#00;
       "GDB_AccessTest".HashData[38] := BYTE#16#00;
       "GDB_AccessTest".HashData[39] := BYTE#16#00;
       "GDB_AccessTest".HashData[40] := BYTE#16#00;
       "GDB_AccessTest".HashData[41] := BYTE#16#00;
       "GDB_AccessTest".HashData[42] := BYTE#16#00;
       "GDB_AccessTest".HashData[43] := BYTE#16#00;
       "GDB_AccessTest".HashData[44] := BYTE#16#00;
       "GDB_AccessTest".HashData[45] := BYTE#16#00;
       "GDB_AccessTest".HashData[46] := BYTE#16#00;
       "GDB_AccessTest".HashData[47] := BYTE#16#00;
       "GDB_AccessTest".HashOk := "FRK_Sha256Pin"(Data := "GDB_AccessTest".HashData, Size := 3, Digest := "GDB_AccessTest".Hash1);
       "GDB_AccessTest".HashData[0] := BYTE#16#00;
       "GDB_AccessTest".HashData[1] := BYTE#16#01;
       "GDB_AccessTest".HashData[2] := BYTE#16#02;
       "GDB_AccessTest".HashData[3] := BYTE#16#03;
       "GDB_AccessTest".HashData[4] := BYTE#16#04;
       "GDB_AccessTest".HashData[5] := BYTE#16#05;
       "GDB_AccessTest".HashData[6] := BYTE#16#06;
       "GDB_AccessTest".HashData[7] := BYTE#16#07;
       "GDB_AccessTest".HashData[8] := BYTE#16#08;
       "GDB_AccessTest".HashData[9] := BYTE#16#09;
       "GDB_AccessTest".HashData[10] := BYTE#16#0A;
       "GDB_AccessTest".HashData[11] := BYTE#16#0B;
       "GDB_AccessTest".HashData[12] := BYTE#16#0C;
       "GDB_AccessTest".HashData[13] := BYTE#16#0D;
       "GDB_AccessTest".HashData[14] := BYTE#16#0E;
       "GDB_AccessTest".HashData[15] := BYTE#16#0F;
       "GDB_AccessTest".HashData[16] := BYTE#16#10;
       "GDB_AccessTest".HashData[17] := BYTE#16#11;
       "GDB_AccessTest".HashData[18] := BYTE#16#12;
       "GDB_AccessTest".HashData[19] := BYTE#16#13;
       "GDB_AccessTest".HashData[20] := BYTE#16#14;
       "GDB_AccessTest".HashData[21] := BYTE#16#15;
       "GDB_AccessTest".HashData[22] := BYTE#16#16;
       "GDB_AccessTest".HashData[23] := BYTE#16#17;
       "GDB_AccessTest".HashData[24] := BYTE#16#18;
       "GDB_AccessTest".HashData[25] := BYTE#16#19;
       "GDB_AccessTest".HashData[26] := BYTE#16#1A;
       "GDB_AccessTest".HashData[27] := BYTE#16#1B;
       "GDB_AccessTest".HashData[28] := BYTE#16#1C;
       "GDB_AccessTest".HashData[29] := BYTE#16#1D;
       "GDB_AccessTest".HashData[30] := BYTE#16#1E;
       "GDB_AccessTest".HashData[31] := BYTE#16#1F;
       "GDB_AccessTest".HashData[32] := BYTE#16#20;
       "GDB_AccessTest".HashData[33] := BYTE#16#21;
       "GDB_AccessTest".HashData[34] := BYTE#16#22;
       "GDB_AccessTest".HashData[35] := BYTE#16#23;
       "GDB_AccessTest".HashData[36] := BYTE#16#24;
       "GDB_AccessTest".HashData[37] := BYTE#16#25;
       "GDB_AccessTest".HashData[38] := BYTE#16#26;
       "GDB_AccessTest".HashData[39] := BYTE#16#27;
       "GDB_AccessTest".HashData[40] := BYTE#16#28;
       "GDB_AccessTest".HashData[41] := BYTE#16#29;
       "GDB_AccessTest".HashData[42] := BYTE#16#2A;
       "GDB_AccessTest".HashData[43] := BYTE#16#2B;
       "GDB_AccessTest".HashData[44] := BYTE#16#2C;
       "GDB_AccessTest".HashData[45] := BYTE#16#2D;
       "GDB_AccessTest".HashData[46] := BYTE#16#2E;
       "GDB_AccessTest".HashData[47] := BYTE#16#2F;
       "GDB_AccessTest".HashOk := "FRK_Sha256Pin"(Data := "GDB_AccessTest".HashData, Size := 32, Digest := "GDB_AccessTest".Hash2);
       "GDB_AccessTest".HashData[0] := BYTE#16#00;
       "GDB_AccessTest".HashData[1] := BYTE#16#01;
       "GDB_AccessTest".HashData[2] := BYTE#16#02;
       "GDB_AccessTest".HashData[3] := BYTE#16#03;
       "GDB_AccessTest".HashData[4] := BYTE#16#04;
       "GDB_AccessTest".HashData[5] := BYTE#16#05;
       "GDB_AccessTest".HashData[6] := BYTE#16#06;
       "GDB_AccessTest".HashData[7] := BYTE#16#07;
       "GDB_AccessTest".HashData[8] := BYTE#16#08;
       "GDB_AccessTest".HashData[9] := BYTE#16#09;
       "GDB_AccessTest".HashData[10] := BYTE#16#0A;
       "GDB_AccessTest".HashData[11] := BYTE#16#0B;
       "GDB_AccessTest".HashData[12] := BYTE#16#0C;
       "GDB_AccessTest".HashData[13] := BYTE#16#0D;
       "GDB_AccessTest".HashData[14] := BYTE#16#0E;
       "GDB_AccessTest".HashData[15] := BYTE#16#0F;
       "GDB_AccessTest".HashData[16] := BYTE#16#10;
       "GDB_AccessTest".HashData[17] := BYTE#16#11;
       "GDB_AccessTest".HashData[18] := BYTE#16#12;
       "GDB_AccessTest".HashData[19] := BYTE#16#13;
       "GDB_AccessTest".HashData[20] := BYTE#16#14;
       "GDB_AccessTest".HashData[21] := BYTE#16#15;
       "GDB_AccessTest".HashData[22] := BYTE#16#16;
       "GDB_AccessTest".HashData[23] := BYTE#16#17;
       "GDB_AccessTest".HashData[24] := BYTE#16#18;
       "GDB_AccessTest".HashData[25] := BYTE#16#19;
       "GDB_AccessTest".HashData[26] := BYTE#16#1A;
       "GDB_AccessTest".HashData[27] := BYTE#16#1B;
       "GDB_AccessTest".HashData[28] := BYTE#16#1C;
       "GDB_AccessTest".HashData[29] := BYTE#16#1D;
       "GDB_AccessTest".HashData[30] := BYTE#16#1E;
       "GDB_AccessTest".HashData[31] := BYTE#16#1F;
       "GDB_AccessTest".HashData[32] := BYTE#16#20;
       "GDB_AccessTest".HashData[33] := BYTE#16#21;
       "GDB_AccessTest".HashData[34] := BYTE#16#22;
       "GDB_AccessTest".HashData[35] := BYTE#16#23;
       "GDB_AccessTest".HashData[36] := BYTE#16#24;
       "GDB_AccessTest".HashData[37] := BYTE#16#25;
       "GDB_AccessTest".HashData[38] := BYTE#16#26;
       "GDB_AccessTest".HashData[39] := BYTE#16#27;
       "GDB_AccessTest".HashData[40] := BYTE#16#28;
       "GDB_AccessTest".HashData[41] := BYTE#16#29;
       "GDB_AccessTest".HashData[42] := BYTE#16#2A;
       "GDB_AccessTest".HashData[43] := BYTE#16#2B;
       "GDB_AccessTest".HashData[44] := BYTE#16#2C;
       "GDB_AccessTest".HashData[45] := BYTE#16#2D;
       "GDB_AccessTest".HashData[46] := BYTE#16#2E;
       "GDB_AccessTest".HashData[47] := BYTE#16#2F;
       "GDB_AccessTest".HashOk := "FRK_Sha256Pin"(Data := "GDB_AccessTest".HashData, Size := 48, Digest := "GDB_AccessTest".Hash3);
       "GDB_RoutingTest".PermitOne := TRUE;
       "GDB_RoutingTest".PermitTwo := TRUE;
       "GDB_RoutingTest".RootManualPermit := TRUE;
       "GDB_RoutingTest".NestedFinish := FALSE;
       "GDB_RoutingTest".InnerFinish := FALSE;
       "GDB_RoutingTest".NestedAccessLock := FALSE;
       #ResultCode := RD_SYS_T(OUT => #StartupStamp);
       IF #ResultCode = 0 THEN
           "GDB_UnitTest".BootStamp := DTL_TO_LDT(#StartupStamp);
       END_IF;
       "GDB_UnitTest".Restarts := "GDB_UnitTest".Restarts + 1;
       "GDB_UnitTest".FinishCycle := FALSE;
       "GDB_UnitTest".Permit := TRUE;
       "GDB_UnitTest".FaultRoot := FALSE;
       "GDB_UnitTest".ExitHold := FALSE;
       "GDB_UnitTest".IssueChild := FALSE;
       "GDB_UnitTest".LockStart := FALSE;
       "GDB_UnitTest".ChildCommand := 2;
       "GDB_UnitTest".Verdict := 1;
       "GDB_UnitTest".Reason := 2003;
       "GDB_UnitTest".CarrierControl := 0;
       "FRK_UnitSetLocalCarrier"(Unit := "StationA".Unit,
                                 Index := 1);
   END_IF;
   "GDB_FraktalHal".Data.StationA.Cell.Clamp.Finish := "GDB_UnitTest".FinishCycle;
   "GDB_FraktalHal".Data.StationA.Cell.Clamp.Permit := "GDB_UnitTest".Permit;
   "GDB_FraktalHal".Data.StationA.Cell.Clamp.ExitHold := "GDB_UnitTest".ExitHold;
   "GDB_FraktalHal".Data.StationA.Cell.Clamp.BackgroundFault := "GDB_UnitTest".FaultRoot;
   "GDB_FraktalHal".Data.StationA.Cell.Clamp.Verdict := "GDB_UnitTest".Verdict;
   "GDB_FraktalHal".Data.StationA.Cell.Clamp.Diag.ReasonCode := "GDB_UnitTest".Reason;
   "GDB_FraktalHal".Data.StationA.Cell.Clamp.Diag.Description := WSTRING#'test.start.permit';
   "GDB_FraktalHal".Data.StationA.Cell.Clamp.Diag.SourcePath := WSTRING#'StationA.Cell.Clamp';
   IF "GDB_UnitTest".IssueChild THEN
       "StationA".Cell.Clamp.Command := "GDB_UnitTest".ChildCommand;
       "StationA".Cell.Clamp.Execute := TRUE;
       "GDB_UnitTest".IssueChild := FALSE;
   END_IF;
   CASE "GDB_UnitTest".CarrierControl OF
       1:
           "FRK_UnitSetLocalCarrier"(Unit := "StationA".Unit,
                                     Index := 1);
       2:
           "FRK_Carriers".Slots[1].Enabled := FALSE;
       3:
           "FRK_Carriers".Slots[1].Context.Uid := 'other';
       ELSE
           "GDB_UnitTest".CarrierControl := 0;
   END_CASE;
   "GDB_UnitTest".CarrierControl := 0;
   "StationA".Cell.Gate.ParCfg.Timeout := T#8s;
   "GDB_FraktalHal".Data.StationA.Cell.Gate.Permit := "GDB_RoutingTest".PermitOne;
   IF "GDB_RoutingTest".PermitTwo THEN
       "GDB_FraktalHal".Data.StationA.Cell.Gate.Sample := 0;
   ELSE
       "GDB_FraktalHal".Data.StationA.Cell.Gate.Sample := 1;
   END_IF;
   "GDB_FraktalHal".Data.StationA.Cell.Gate.Diag.ReasonCode := 2002;
   "GDB_FraktalHal".Data.StationA.Cell.Gate.Diag.Description := WSTRING#'test.manual.first';
   "GDB_FraktalHal".Data.StationA.Cell.Gate.LaterDiag.ReasonCode := 2003;
   "GDB_FraktalHal".Data.StationA.Cell.Gate.LaterDiag.Description := WSTRING#'test.manual.second';
   "GDB_FraktalHal".Data.StationA.Satellite.Cell.Clamp.Permit := "GDB_RoutingTest".RootManualPermit;
   "GDB_FraktalHal".Data.StationA.Satellite.Cell.Clamp.Diag.SourcePath := WSTRING#'StationA.Satellite.Cell.Clamp';
   "GDB_FraktalHal".Data.StationA.Satellite.Cell.Clamp.Diag.Description := WSTRING#'test.nested.permit';
   "GDB_FraktalHal".Data.StationA.Satellite.Cell.Clamp.Diag.ReasonCode := 2002;
   "GDB_FraktalHal".Data.StationA.Satellite.Inner.Cell.Clamp.Permit := TRUE;
   "GDB_FraktalHal".Data.StationA.Satellite.Cell.Clamp.Finish := "GDB_RoutingTest".NestedFinish;
   "GDB_FraktalHal".Data.StationA.Satellite.Inner.Cell.Clamp.Finish := "GDB_RoutingTest".InnerFinish;
   IF "GDB_RoutingTest".NestedAccessLock THEN
       "StationA".Satellite.Access.Policy.Required[5] := 4;
   ELSE
       "StationA".Satellite.Access.Policy.Required[5] := 0;
   END_IF;
   IF "GDB_RoutingTest".LocalPulse THEN
       "GDB_RoutingTest".LocalRequest.Kind := "GDB_RoutingTest".LocalKind;
       "GDB_RoutingTest".LocalRequest.IntValue := "GDB_RoutingTest".LocalValue;
       "FRK_UnitOperation"(Core := "StationA".Satellite.Core,
                           Unit := "StationA".Satellite.Unit,
                           Status := "StationA".Satellite.Status,
                           Policy := "StationA".Satellite.ModePolicy,
                           Access := "StationA".Satellite.Access,
                           Supported := "StationA".Satellite.SupportedModesPublished,
                           Request := "GDB_RoutingTest".LocalRequest,
                           Response := "FRK_UnitScratch".Response,
                           Trusted := FALSE);
       "GDB_RoutingTest".LocalAccepted := "FRK_UnitScratch".Response.Accepted;
       "GDB_RoutingTest".LocalFirstKind := -1;
       IF "FRK_UnitScratch".Response.Report.Count > 0 THEN
           "GDB_RoutingTest".LocalFirstKind := "FRK_UnitScratch".Response.Report.Reasons[1].Kind;
       END_IF;
       "GDB_RoutingTest".LocalPulse := FALSE;
   END_IF;
   "StationA".Access.ProviderEnabled := NOT "GDB_AccessTest".ProviderOff;
   "StationB".Access.ProviderEnabled := NOT "GDB_AccessTest".ProviderOff;
   "GDB_FraktalMain"(Startup := #Initial_Call);
   "GDB_RoutingTest".ManExecute := "StationA".Cell.Gate.Execute;
   "GDB_RoutingTest".ManStarts := "StationA".Cell.Gate.Device.StartCount;
   "GDB_UnitTest".Scans := "GDB_UnitTest".Scans + 1;
   "GDB_UnitTest".ChildExecute := "StationA".Cell.Clamp.Execute;
   "GDB_UnitTest".ChildState := "StationA".Cell.Clamp.Core.Exec;
   "GDB_UnitTest".CarrierWrites := "FRK_Carriers".Slots[1].Writes;
   "GDB_UnitTest".CarrierSerial := "FRK_Carriers".Slots[1].Serial;
   "GDB_UnitTest".WrittenUid := "FRK_Carriers".Slots[1].Written.Uid;
   "GDB_UnitTest".WrittenVerdict := "FRK_Carriers".Slots[1].Written.Result.Verdict;
   IF "StationA".HistoryHead > 0 AND "StationA".HistoryHead <= 16 THEN
       "GDB_UnitTest".LastEvent := "StationA".History["StationA".HistoryHead].ReasonCode;
   END_IF;
   "GDB_UnitTest".SecretCleared := "StationA".HmiRequest.Secret = '';
   "GDB_UnitTest".SnapshotSecretCleared := "StationA".Unit.Request.Secret = '';
   IF "StationA".Access.LoginBusy AND ("GDB_AccessTest".CancelOnLogin OR "GDB_AccessTest".SupersedeOnLogin) THEN
       "GDB_AccessTest".InterruptedBusy := TRUE;
       IF "GDB_AccessTest".CancelOnLogin THEN
           "GDB_AccessTest".InterruptRequest.Kind := 2;
           "FRK_UnitOperation"(Core := "StationA".Core,
                               Unit := "StationA".Unit,
                               Status := "StationA".Status,
                               Policy := "StationA".ModePolicy,
                               Access := "StationA".Access,
                               Supported := "StationA".SupportedModesPublished,
                               Request := "GDB_AccessTest".InterruptRequest,
                               Response := "FRK_UnitScratch".Response,
                               Trusted := FALSE);
       ELSE
           "GDB_AccessTest".SupersededSequence := "FRK_AccessNext"(Previous := "StationA".Access.LoginSequence);
           "FRK_AccessLogin"(Access := "StationA".Access,
                             User := 'unknown',
                             Secret := 'wrong',
                             Sequence := "GDB_AccessTest".SupersededSequence);
       END_IF;
       "GDB_AccessTest".CancelOnLogin := FALSE;
       "GDB_AccessTest".SupersedeOnLogin := FALSE;
   END_IF;
END_ORGANIZATION_BLOCK

FUNCTION_BLOCK "FB_FraktalMain"   // FB6, SCL
{ S7_Optimized_Access := 'TRUE' }
VERSION : 0.1
// stored: AutoNumber true, IsIECCheckEnabled false, IsRetainMemResEnabled false, MemoryReserve 100, SetENOAutomatically false, UDAEnableTagReadback false
   VAR_INPUT
      Startup { ExternalAccessible := 'False'; ExternalVisible := 'False'; ExternalWritable := 'False'} : Bool;
   END_VAR
BEGIN

   IF #Startup THEN
       "FRK_Registry".Count := 0;
       "FRK_Registry".Fault := FALSE;
   END_IF;
   "FRK_ClockTick"();
   "StationA"(ParentIndex := 0,
              Startup := #Startup,
              Hal := "GDB_FraktalHal".Data.StationA);
   "StationB"(ParentIndex := 0,
              Startup := #Startup,
              Hal := "GDB_FraktalHal".Data.StationB);
END_FUNCTION_BLOCK

FUNCTION_BLOCK "FB_DeclarationUnit"   // FB5, SCL
{ S7_Optimized_Access := 'TRUE' }
VERSION : 0.1
// Generated frame v0.6; change the declaration, then regenerate.
// stored: AutoNumber true, IsIECCheckEnabled false, IsRetainMemResEnabled false, MemoryReserve 100, SetENOAutomatically false, UDAEnableTagReadback false
   VAR_INPUT
      Execute { ExternalWritable := 'False'} : Bool;
      Abort { ExternalWritable := 'False'} : Bool;
      Command { ExternalWritable := 'False'} : DInt;
      ParCfg { ExternalWritable := 'False'} : "ST_DeclarationParCfg";
      ParCmd { ExternalWritable := 'False'} : "ST_DeclarationParCmd";
      ParentIndex { ExternalAccessible := 'False'; ExternalVisible := 'False'; ExternalWritable := 'False'} : DInt;
      Startup { ExternalAccessible := 'False'; ExternalVisible := 'False'; ExternalWritable := 'False'} : Bool;
   END_VAR
   VAR_OUTPUT
      Busy { ExternalWritable := 'False'} : Bool;
      Done { ExternalWritable := 'False'} : Bool;
      Error { ExternalWritable := 'False'} : Bool;
      Aborted { ExternalWritable := 'False'} : Bool;
      Held { ExternalWritable := 'False'} : Bool;
      ErrorID { ExternalWritable := 'False'} : DWord;
      Timing { ExternalWritable := 'False'} : "ST_ModuleTiming";
      OutCmd { ExternalWritable := 'False'} : "ST_DeclarationOutCmd";
      OutImm { ExternalWritable := 'False'} : "ST_UnitProbeImm";
   END_VAR
   VAR_IN_OUT
      Hal : "ST_DeclarationUnitHal";
   END_VAR
   VAR
      Status { ExternalWritable := 'False'; S7_SetPoint := 'True'} : "ST_ModuleStatus";
      Core { ExternalAccessible := 'False'; ExternalVisible := 'False'; ExternalWritable := 'False'; S7_SetPoint := 'True'} : "FRK_Core";
      LatchedParCmd { ExternalAccessible := 'False'; ExternalVisible := 'False'; ExternalWritable := 'False'; S7_SetPoint := 'True'} : "ST_DeclarationParCmd";
      Device { ExternalAccessible := 'False'; ExternalVisible := 'False'; ExternalWritable := 'False'; S7_SetPoint := 'True'} : "ST_UnitProbeDevice";
      Unit { ExternalAccessible := 'False'; ExternalVisible := 'False'; ExternalWritable := 'False'; S7_SetPoint := 'True'} : "FRK_Unit";
      HmiRequest { S7_SetPoint := 'True'} : "ST_HmiRequest";
      ModePolicy { ExternalAccessible := 'False'; ExternalVisible := 'False'; ExternalWritable := 'False'; S7_SetPoint := 'True'} : Array[0..6] of "ST_ModePolicy";
      Access { ExternalWritable := 'False'; S7_SetPoint := 'True'} : "FRK_Access";
      HmiResponse { ExternalWritable := 'False'; S7_SetPoint := 'True'} : "ST_HmiResponse";
      ConfigRev { ExternalWritable := 'False'} : UDInt;
      ConfigCursor { ExternalAccessible := 'False'; ExternalVisible := 'False'; ExternalWritable := 'False'; S7_SetPoint := 'True'} : "FRK_ConfigCursor";
      Part { ExternalWritable := 'False'; S7_SetPoint := 'True'} : "ST_PartContext";
      History { ExternalWritable := 'False'; S7_SetPoint := 'True'} : Array[1..16] of "ST_Diagnostic";
      HistoryHead { ExternalWritable := 'False'} : Int;
      ModeActivePublished { ExternalWritable := 'False'} : DInt;
      RunningPublished { ExternalWritable := 'False'} : Bool;
      StopPendingPublished { ExternalWritable := 'False'} : Bool;
      SupportedModesPublished { ExternalWritable := 'False'} : Array[0..6] of Bool;
      GoodCount { ExternalWritable := 'False'} : UDInt;
      NokCount { ExternalWritable := 'False'} : UDInt;
      ReworkCount { ExternalWritable := 'False'} : UDInt;
      NokReason { ExternalWritable := 'False'} : DInt;
      Cell { ExternalWritable := 'False'; S7_SetPoint := 'True'} : "FB_DeclarationCell";
      Satellite { ExternalWritable := 'False'; S7_SetPoint := 'True'} : "FB_SatelliteUnit";
   END_VAR
   VAR_TEMP
      InstancePath : WString[254];
      RouteMatched : Bool;
      ManualMatched : Bool;
   END_VAR
   VAR CONSTANT
      EXEC_READY : DInt := 0;
      MODULE_TIER : DInt := 1;
   END_VAR
BEGIN

   // ---- GENERATED: setup
   IF #Startup OR NOT #Core.Named THEN
       #InstancePath := GetInstancePath(size := 0);
       "FRK_SetIdentity"(Core := #Core,
                         Status := #Status,
                         InstancePath := #InstancePath,
                         ModuleType := 1,
                         TypeId := 1,
                         Capabilities := DWORD#16#00000000,
                         ParentIndex := #ParentIndex,
                         TypeKey := 'Fraktal.Declaration.Unit');
   END_IF;
   IF #Startup OR #ConfigRev = 0 THEN
       #ConfigRev := "FRK_ConfigRevision"(Previous := #ConfigRev);
   END_IF;
   #SupportedModesPublished[0] := TRUE;
   #SupportedModesPublished[1] := TRUE;
   #SupportedModesPublished[2] := TRUE;
   #SupportedModesPublished[3] := TRUE;
   #SupportedModesPublished[4] := FALSE;
   #SupportedModesPublished[5] := FALSE;
   #SupportedModesPublished[6] := FALSE;
   "FRK_UnitPrepare"(Core := #Core,
                     Unit := #Unit,
                     Policy := #ModePolicy,
                     Request := #HmiRequest,
                     Response := #HmiResponse,
                     Startup := #Startup,
                     InitialMode := 1);
   "FRK_AccessCyclic"(Access := #Access,
                      Startup := #Startup,
                      SourcePath := STRING_TO_WSTRING(#Status.Name),
                      History := #History,
                      Head := #HistoryHead,
                      Revision := #ConfigRev);
   "FRK_UnitMailbox"(Core := #Core,
                     Unit := #Unit,
                     Status := #Status,
                     Policy := #ModePolicy,
                     Access := #Access,
                     Request := #HmiRequest,
                     Response := #HmiResponse,
                     Supported := #SupportedModesPublished);
   // ---- GENERATED: begin
   "FRK_Begin"(Core := #Core,
               Status := #Status,
               Execute := #Unit.RunReq,
               Abort := (#Abort OR #Unit.AbortReq),
               Command := 1);
   IF #Core.EvCommandStart THEN
       #LatchedParCmd := #ParCmd;
       CASE #Core.Command OF
           1:
               "FRK_UnitRunStart"(Core := #Core,
                                  Status := #Status,
                                  Timeout := #ParCfg.Timeout,
                                  Label := 'Run');
           ELSE
               "FRK_Start"(Core := #Core,
                           Status := #Status,
                           Supported := FALSE,
                           Timeout := T#0ms,
                           Label := '');
       END_CASE;
   END_IF;
   IF #Core.EvCommandStart THEN
       // ---- AUTHORED: CommandStart
       #Device.Received := "FRK_PartReceived"(Core := #Core, Unit := #Unit, Status := #Status, Part := #Part, History := #History, Head := #HistoryHead);
       IF #Device.Received THEN
           "FRK_PartStarted"(Unit := #Unit,
                             Status := #Status,
                             Part := #Part,
                             History := #History,
                             Head := #HistoryHead);
       END_IF;
       // ---- GENERATED: reaction end
   END_IF;
   // ---- AUTHORED: cyclic management
   IF #Hal.Cell.Clamp.BackgroundFault THEN
       "FRK_Fault"(Core := #Core,
                   Status := #Status,
                   ReasonCode := 2901,
                   Description := WSTRING#'test.unit.condition');
   END_IF;
   // ---- GENERATED: end management
   "FRK_Release_DeclarationUnit"(Unit := #Unit,
                                 Hal := #Hal);
   "FRK_UnitConsume"(Core := #Core,
                     Unit := #Unit,
                     Status := #Status,
                     Policy := #ModePolicy,
                     Access := #Access,
                     Response := #HmiResponse,
                     Supported := #SupportedModesPublished);
   "FRK_UnitMode"(Core := #Core,
                  Unit := #Unit);
   IF #Core.EvModeExit THEN
       // ---- AUTHORED: ModeExit
       #Device.ExitCalls := #Device.ExitCalls + 1;
       IF #Hal.Cell.Clamp.ExitHold THEN
           #Core.HookResult := 1;
       ELSE
           #Core.HookResult := 0;
       END_IF;
       // ---- GENERATED: reaction end
   END_IF;
   "FRK_UnitModeResolve"(Core := #Core,
                         Unit := #Unit,
                         Status := #Status,
                         Policy := #ModePolicy,
                         Timeout := #ParCfg.Timeout);
   IF #Core.EvModeChanged THEN
       // ---- AUTHORED: ModeChanged
       #Device.Changes := #Device.Changes + 1;
       // ---- GENERATED: reaction end
   END_IF;
   "FRK_UnitFollow"(Core := #Core,
                    Unit := #Unit,
                    Status := #Status,
                    Policy := #ModePolicy,
                    Access := #Access,
                    Supported := #SupportedModesPublished);
   IF #Unit.RequestPending AND (#Unit.Request.Kind = 11 OR #Unit.Request.Kind = 16) THEN
       #ManualMatched := FALSE;
       #RouteMatched := "FRK_Route_DeclarationCell"(Module := #Cell, Hal := #Hal.Cell, Request := #Unit.Request, Report := #HmiResponse.Report);
       #ManualMatched := #ManualMatched OR #RouteMatched;
       #RouteMatched := "FRK_Route_SatelliteUnit"(Module := #Satellite, Hal := #Hal.Satellite, Request := #Unit.Request, Report := #HmiResponse.Report);
       #ManualMatched := #ManualMatched OR #RouteMatched;
       IF NOT #ManualMatched THEN
           "FRK_ReleaseReason"(Report := #HmiResponse.Report,
                               Description := WSTRING#'std.error.unsupportedHmiRequest',
                               Reason := 2008,
                               Path := #Unit.Request.TargetPath,
                               Kind := 4);
       END_IF;
       #HmiResponse.Accepted := #Unit.Request.Kind = 16 OR #HmiResponse.Report.Released;
       IF #Unit.Request.Kind = 11 THEN
           IF #HmiResponse.Accepted THEN
               #HmiResponse.Diagnostic := WSTRING#'std.audit.manualCommandAccepted';
           ELSE
               #HmiResponse.Diagnostic := WSTRING#'std.audit.manualCommandRejected';
           END_IF;
       END_IF;
   END_IF;
   IF #Unit.EvReset THEN
       // ---- AUTHORED: OperatorReset
       #Device.Resets := #Device.Resets + 1;
       // ---- GENERATED: reset reaction end
   END_IF;
   IF #Core.ReleasePending OR #Unit.ReleaseChildren THEN
       "FRK_ReleaseCommand"(Core := #Cell.Core,
                            Execute := #Cell.Execute);
       "FRK_ReleaseCommand"(Core := #Satellite.Core,
                            Execute := #Satellite.Execute);
   END_IF;
   // ---- GENERATED: child call
   #Cell(ParentIndex := #Core.RegIndex,
         Startup := #Startup,
         Hal := #Hal.Cell);
   "FRK_ManualFinish"(Core := #Cell.Core,
                      Execute := #Cell.Execute,
                      ManualOwned := #Cell.ManualOwned);
   "FRK_UnitCascade"(ParentUnit := #Unit,
                     Core := #Satellite.Core,
                     Unit := #Satellite.Unit,
                     Status := #Satellite.Status,
                     Policy := #Satellite.ModePolicy,
                     Access := #Satellite.Access,
                     Supported := #Satellite.SupportedModesPublished,
                     History := #History,
                     Head := #HistoryHead);
   // ---- GENERATED: child call
   #Satellite(ParentIndex := #Core.RegIndex,
              Startup := #Startup,
              Hal := #Hal.Satellite);
   #Unit.CascadePending := FALSE;
   IF #Unit.RequestPending AND #Unit.Request.Kind = 23 THEN
       #HmiResponse.Accepted := FALSE;
       #HmiResponse.Report.Count := 0;
       #HmiResponse.Report.Released := TRUE;
       #HmiResponse.Diagnostic := WSTRING#'';
       "FRK_ConfigBegin"(Cursor := #ConfigCursor,
                         Page := #HmiResponse.ConfigPage,
                         PageIndex := #Unit.Request.IntValue,
                         Revision := #ConfigRev);
       IF #Unit.Request.DurationMs <> 0 THEN
           #HmiResponse.Diagnostic := WSTRING#'std.error.modelNotAvailable';
       ELSIF #Unit.Request.IntValue < 0 OR #Unit.Request.IntValue > 32767 THEN
           #HmiResponse.Diagnostic := WSTRING#'std.error.hmiRequestRejected';
       ELSE
           "FRK_ConfigUnit"(Scope := #Status.Name,
                            Policy := #ModePolicy,
                            ReadLevel := #Access.Policy.Required[0],
                            Readable := #Access.CurrentLevel >= #Access.Policy.Required[0],
                            Cursor := #ConfigCursor,
                            Page := #HmiResponse.ConfigPage);
           "FRK_Config_DeclarationCell"(Module := #Cell,
                                        ReadLevel := #Access.Policy.Required[0],
                                        Readable := #Access.CurrentLevel >= #Access.Policy.Required[0],
                                        Cursor := #ConfigCursor,
                                        Page := #HmiResponse.ConfigPage);
           "FRK_Config_SatelliteUnit"(Module := #Satellite,
                                      ReadLevel := #Access.Policy.Required[0],
                                      Readable := #Access.CurrentLevel >= #Access.Policy.Required[0],
                                      Cursor := #ConfigCursor,
                                      Page := #HmiResponse.ConfigPage);
           "FRK_ConfigFinish"(Cursor := #ConfigCursor,
                              Page := #HmiResponse.ConfigPage);
           #HmiResponse.Accepted := TRUE;
       END_IF;
   END_IF;
   "FRK_RouteAbort"(Core := #Core,
                    Abort := (#Abort OR #Unit.AbortReq));
   IF #Core.EvAbort THEN
       "FRK_PartAborted"(Core := #Core,
                         Unit := #Unit,
                         Status := #Status,
                         Part := #Part,
                         History := #History,
                         Head := #HistoryHead);
   END_IF;
   IF #Core.Dispatch AND #Core.RegIndex > 0 AND NOT "FRK_Registry".Fault THEN
       // ---- AUTHORED: dispatch
       IF #Hal.Cell.Clamp.Finish THEN
           #Device.Processed := FALSE;
           IF #Unit.CarrierIndex = 0 THEN
               #Device.Processed := TRUE;
           ELSE
               #Device.Processed := "FRK_PartProcessed"(Core := #Core, Unit := #Unit, Status := #Status, Part := #Part, History := #History, Head := #HistoryHead, Verdict := #Hal.Cell.Clamp.Verdict, Reason := #Hal.Cell.Clamp.Diag.ReasonCode);
           END_IF;
           IF #Device.Processed THEN
               #Device.Cycles := #Device.Cycles + 1;
               IF #Unit.StopReq THEN
                   "FRK_Complete"(Core := #Core,
                                  Status := #Status);
               ELSE
                   #Device.Received := "FRK_PartReceived"(Core := #Core, Unit := #Unit, Status := #Status, Part := #Part, History := #History, Head := #HistoryHead);
                   IF #Device.Received THEN
                       "FRK_PartStarted"(Unit := #Unit,
                                         Status := #Status,
                                         Part := #Part,
                                         History := #History,
                                         Head := #HistoryHead);
                   END_IF;
               END_IF;
           END_IF;
       END_IF;
       // ---- GENERATED: end dispatch
   END_IF;
   "FRK_End"(Core := #Core,
             Status := #Status,
             Busy => #Busy,
             Done => #Done,
             Error => #Error,
             Aborted => #Aborted,
             Held => #Held,
             ErrorID => #ErrorID,
             Timing => #Timing);
   "FRK_AccessFinish"(Access := #Access,
                      Unit := #Unit,
                      Response := #HmiResponse,
                      SourcePath := STRING_TO_WSTRING(#Status.Name),
                      History := #History,
                      Head := #HistoryHead,
                      Revision := #ConfigRev);
   "FRK_UnitFinish"(Core := #Core,
                    Unit := #Unit,
                    Response := #HmiResponse,
                    Status := #Status,
                    Part := #Part,
                    History := #History,
                    Head := #HistoryHead);
   #ModeActivePublished := #Unit.Mode;
   #RunningPublished := #Core.Exec = 1;
   #StopPendingPublished := #Unit.StopReq AND #Core.Exec = 1;
   #GoodCount := #Unit.Good;
   #NokCount := #Unit.Nok;
   #ReworkCount := #Unit.Rework;
   #NokReason := #Unit.NokReason;
   // ---- AUTHORED: unconditional cyclic/derived data
   #OutImm.Cycles := #Device.Cycles;
   #OutImm.ExitCalls := #Device.ExitCalls;
   #OutImm.Changes := #Device.Changes;
   #OutImm.Resets := #Device.Resets;
   // ---- GENERATED: frame end
END_FUNCTION_BLOCK

FUNCTION_BLOCK "FB_DeclarationCell"   // FB2, SCL
{ S7_Optimized_Access := 'TRUE' }
VERSION : 0.1
// Generated frame v0.6; change the declaration, then regenerate.
// stored: AutoNumber true, IsIECCheckEnabled false, IsRetainMemResEnabled false, MemoryReserve 100, SetENOAutomatically false, UDAEnableTagReadback false
   VAR_INPUT
      Execute { ExternalWritable := 'False'} : Bool;
      Abort { ExternalWritable := 'False'} : Bool;
      Command { ExternalWritable := 'False'} : DInt;
      ParCfg { ExternalWritable := 'False'} : "ST_DeclarationParCfg";
      ParCmd { ExternalWritable := 'False'} : "ST_DeclarationParCmd";
      ParentIndex { ExternalAccessible := 'False'; ExternalVisible := 'False'; ExternalWritable := 'False'} : DInt;
      Startup { ExternalAccessible := 'False'; ExternalVisible := 'False'; ExternalWritable := 'False'} : Bool;
   END_VAR
   VAR_OUTPUT
      Busy { ExternalWritable := 'False'} : Bool;
      Done { ExternalWritable := 'False'} : Bool;
      Error { ExternalWritable := 'False'} : Bool;
      Aborted { ExternalWritable := 'False'} : Bool;
      Held { ExternalWritable := 'False'} : Bool;
      ErrorID { ExternalWritable := 'False'} : DWord;
      Timing { ExternalWritable := 'False'} : "ST_ModuleTiming";
      OutCmd { ExternalWritable := 'False'} : "ST_DeclarationOutCmd";
      OutImm { ExternalWritable := 'False'} : "ST_DeclarationOutImm";
   END_VAR
   VAR_IN_OUT
      Hal : "ST_DeclarationCellHal";
   END_VAR
   VAR
      Status { ExternalWritable := 'False'; S7_SetPoint := 'True'} : "ST_ModuleStatus";
      Core { ExternalAccessible := 'False'; ExternalVisible := 'False'; ExternalWritable := 'False'; S7_SetPoint := 'True'} : "FRK_Core";
      LatchedParCmd { ExternalAccessible := 'False'; ExternalVisible := 'False'; ExternalWritable := 'False'; S7_SetPoint := 'True'} : "ST_DeclarationParCmd";
      Device { ExternalAccessible := 'False'; ExternalVisible := 'False'; ExternalWritable := 'False'; S7_SetPoint := 'True'} : "ST_DeclarationOutImm";
      Catalog { ExternalAccessible := 'False'; ExternalVisible := 'False'; ExternalWritable := 'False'; S7_SetPoint := 'True'} : Array[1..12] of "ST_CommandInfo";
      CatalogCount { ExternalAccessible := 'False'; ExternalVisible := 'False'; ExternalWritable := 'False'} : Int;
      ManConditions { ExternalAccessible := 'False'; ExternalVisible := 'False'; ExternalWritable := 'False'; S7_SetPoint := 'True'} : Array[1..16] of "FRK_ManualConditionRow";
      ManualOwned { ExternalAccessible := 'False'; ExternalVisible := 'False'; ExternalWritable := 'False'} : Bool;
      Clamp { ExternalWritable := 'False'; S7_SetPoint := 'True'} : "FB_DeclarationCylinder";
      Gate { ExternalWritable := 'False'; S7_SetPoint := 'True'} : "FB_DeclarationCylinder";
   END_VAR
   VAR_TEMP
      InstancePath : WString[254];
   END_VAR
   VAR CONSTANT
      EXEC_READY : DInt := 0;
      MODULE_TIER : DInt := 2;
   END_VAR
BEGIN

   // ---- GENERATED: setup
   IF #Startup OR NOT #Core.Named THEN
       #InstancePath := GetInstancePath(size := 0);
       "FRK_SetIdentity"(Core := #Core,
                         Status := #Status,
                         InstancePath := #InstancePath,
                         ModuleType := 2,
                         TypeId := 2,
                         Capabilities := DWORD#16#00000000,
                         ParentIndex := #ParentIndex,
                         TypeKey := 'Fraktal.Declaration.Cell');
       #CatalogCount := 7;
       #Catalog[1].Value := 1;
       #Catalog[1].Label := 'Finish';
       #Catalog[1].Style := 0;
       #Catalog[2].Value := 2;
       #Catalog[2].Label := 'Wait';
       #Catalog[2].Style := 0;
       #Catalog[3].Value := 3;
       #Catalog[3].Label := 'Hold';
       #Catalog[3].Style := 0;
       #Catalog[4].Value := 4;
       #Catalog[4].Label := 'Fault';
       #Catalog[4].Style := 0;
       #Catalog[5].Value := 5;
       #Catalog[5].Label := 'Pending';
       #Catalog[5].Style := 0;
       #Catalog[6].Value := 6;
       #Catalog[6].Label := 'Instant';
       #Catalog[6].Style := 0;
       #Catalog[7].Value := 7;
       #Catalog[7].Label := 'Adopt';
       #Catalog[7].Style := 0;
   END_IF;
   // ---- GENERATED: begin
   "FRK_Begin"(Core := #Core,
               Status := #Status,
               Execute := #Execute,
               Abort := #Abort,
               Command := #Command);
   IF #Core.EvInit THEN
       // ---- AUTHORED: Init
       #Device.InitCount := #Device.InitCount + 1;
       // ---- GENERATED: reaction end
   END_IF;
   IF #Core.EvCommandStart THEN
       #LatchedParCmd := #ParCmd;
       CASE #Core.Command OF
           1:
               "FRK_Start"(Core := #Core,
                           Status := #Status,
                           Supported := TRUE,
                           Timeout := #ParCfg.Timeout,
                           Label := 'Finish');
           2:
               "FRK_Start"(Core := #Core,
                           Status := #Status,
                           Supported := TRUE,
                           Timeout := #ParCfg.Timeout,
                           Label := 'Wait');
           3:
               "FRK_Start"(Core := #Core,
                           Status := #Status,
                           Supported := TRUE,
                           Timeout := #ParCfg.Timeout,
                           Label := 'Hold');
           4:
               "FRK_Start"(Core := #Core,
                           Status := #Status,
                           Supported := TRUE,
                           Timeout := #ParCfg.Timeout,
                           Label := 'Fault');
           5:
               "FRK_Start"(Core := #Core,
                           Status := #Status,
                           Supported := TRUE,
                           Timeout := #ParCfg.Timeout,
                           Label := 'Pending');
           6:
               "FRK_Start"(Core := #Core,
                           Status := #Status,
                           Supported := TRUE,
                           Timeout := #ParCfg.Timeout,
                           Label := 'Instant');
           7:
               "FRK_Start"(Core := #Core,
                           Status := #Status,
                           Supported := TRUE,
                           Timeout := #ParCfg.Timeout,
                           Label := 'Adopt');
           ELSE
               "FRK_Start"(Core := #Core,
                           Status := #Status,
                           Supported := FALSE,
                           Timeout := T#0ms,
                           Label := '');
       END_CASE;
   END_IF;
   IF #Core.EvCommandStart THEN
       // ---- AUTHORED: CommandStart
       #Device.StartCount := #Device.StartCount + 1;
       #Device.Ordered := #Device.InitCount = 1;
       // ---- GENERATED: reaction end
   END_IF;
   IF #Core.ReleasePending THEN
       "FRK_ReleaseCommand"(Core := #Clamp.Core,
                            Execute := #Clamp.Execute);
       "FRK_ReleaseCommand"(Core := #Gate.Core,
                            Execute := #Gate.Execute);
   END_IF;
   // ---- GENERATED: child call
   #Clamp(ParentIndex := #Core.RegIndex,
          Startup := #Startup,
          Hal := #Hal.Clamp);
   "FRK_ManualFinish"(Core := #Clamp.Core,
                      Execute := #Clamp.Execute,
                      ManualOwned := #Clamp.ManualOwned);
   // ---- GENERATED: child call
   #Gate(ParentIndex := #Core.RegIndex,
         Startup := #Startup,
         Hal := #Hal.Gate);
   "FRK_ManualFinish"(Core := #Gate.Core,
                      Execute := #Gate.Execute,
                      ManualOwned := #Gate.ManualOwned);
   "FRK_RouteAbort"(Core := #Core,
                    Abort := #Abort);
   "FRK_End"(Core := #Core,
             Status := #Status,
             Busy => #Busy,
             Done => #Done,
             Error => #Error,
             Aborted => #Aborted,
             Held => #Held,
             ErrorID => #ErrorID,
             Timing => #Timing);
   // ---- AUTHORED: unconditional cyclic/derived data
   #Device.Sample := #Device.Sample + 1;
   #OutImm := #Device;
   // ---- GENERATED: frame end
END_FUNCTION_BLOCK

FUNCTION_BLOCK "FB_DeclarationCylinder"   // FB1, SCL
{ S7_Optimized_Access := 'TRUE' }
VERSION : 0.1
// Generated frame v0.6; change the declaration, then regenerate.
// stored: AutoNumber true, IsIECCheckEnabled false, IsRetainMemResEnabled false, MemoryReserve 100, SetENOAutomatically false, UDAEnableTagReadback false
   VAR_INPUT
      Execute { ExternalWritable := 'False'} : Bool;
      Abort { ExternalWritable := 'False'} : Bool;
      Command { ExternalWritable := 'False'} : DInt;
      ParCfg { ExternalWritable := 'False'} : "ST_DeclarationParCfg";
      ParCmd { ExternalWritable := 'False'} : "ST_DeclarationParCmd";
      ParentIndex { ExternalAccessible := 'False'; ExternalVisible := 'False'; ExternalWritable := 'False'} : DInt;
      Startup { ExternalAccessible := 'False'; ExternalVisible := 'False'; ExternalWritable := 'False'} : Bool;
   END_VAR
   VAR_OUTPUT
      Busy { ExternalWritable := 'False'} : Bool;
      Done { ExternalWritable := 'False'} : Bool;
      Error { ExternalWritable := 'False'} : Bool;
      Aborted { ExternalWritable := 'False'} : Bool;
      Held { ExternalWritable := 'False'} : Bool;
      ErrorID { ExternalWritable := 'False'} : DWord;
      Timing { ExternalWritable := 'False'} : "ST_ModuleTiming";
      OutCmd { ExternalWritable := 'False'} : "ST_DeclarationOutCmd";
      OutImm { ExternalWritable := 'False'} : "ST_DeclarationOutImm";
   END_VAR
   VAR_IN_OUT
      Hal : "ST_DeclarationLeafHal";
   END_VAR
   VAR
      Status { ExternalWritable := 'False'; S7_SetPoint := 'True'} : "ST_ModuleStatus";
      Core { ExternalAccessible := 'False'; ExternalVisible := 'False'; ExternalWritable := 'False'; S7_SetPoint := 'True'} : "FRK_Core";
      LatchedParCmd { ExternalAccessible := 'False'; ExternalVisible := 'False'; ExternalWritable := 'False'; S7_SetPoint := 'True'} : "ST_DeclarationParCmd";
      Device { ExternalAccessible := 'False'; ExternalVisible := 'False'; ExternalWritable := 'False'; S7_SetPoint := 'True'} : "ST_DeclarationOutImm";
      Catalog { ExternalAccessible := 'False'; ExternalVisible := 'False'; ExternalWritable := 'False'; S7_SetPoint := 'True'} : Array[1..12] of "ST_CommandInfo";
      CatalogCount { ExternalAccessible := 'False'; ExternalVisible := 'False'; ExternalWritable := 'False'} : Int;
      ManConditions { ExternalAccessible := 'False'; ExternalVisible := 'False'; ExternalWritable := 'False'; S7_SetPoint := 'True'} : Array[1..16] of "FRK_ManualConditionRow";
      ManualOwned { ExternalAccessible := 'False'; ExternalVisible := 'False'; ExternalWritable := 'False'} : Bool;
   END_VAR
   VAR_TEMP
      InstancePath : WString[254];
   END_VAR
   VAR CONSTANT
      EXEC_READY : DInt := 0;
      MODULE_TIER : DInt := 3;
   END_VAR
BEGIN

   // ---- GENERATED: setup
   IF #Startup OR NOT #Core.Named THEN
       #InstancePath := GetInstancePath(size := 0);
       "FRK_SetIdentity"(Core := #Core,
                         Status := #Status,
                         InstancePath := #InstancePath,
                         ModuleType := 3,
                         TypeId := 3,
                         Capabilities := DWORD#16#00000000,
                         ParentIndex := #ParentIndex,
                         TypeKey := 'Fraktal.Declaration.Cylinder');
       #CatalogCount := 7;
       #Catalog[1].Value := 1;
       #Catalog[1].Label := 'Finish';
       #Catalog[1].Style := 0;
       #Catalog[2].Value := 2;
       #Catalog[2].Label := 'Wait';
       #Catalog[2].Style := 0;
       #Catalog[3].Value := 3;
       #Catalog[3].Label := 'Hold';
       #Catalog[3].Style := 0;
       #Catalog[4].Value := 4;
       #Catalog[4].Label := 'Fault';
       #Catalog[4].Style := 0;
       #Catalog[5].Value := 5;
       #Catalog[5].Label := 'Pending';
       #Catalog[5].Style := 0;
       #Catalog[6].Value := 6;
       #Catalog[6].Label := 'Instant';
       #Catalog[6].Style := 0;
       #Catalog[7].Value := 7;
       #Catalog[7].Label := 'Adopt';
       #Catalog[7].Style := 0;
   END_IF;
   // ---- GENERATED: begin
   "FRK_Begin"(Core := #Core,
               Status := #Status,
               Execute := #Execute,
               Abort := #Abort,
               Command := #Command);
   IF #Core.EvInit THEN
       // ---- AUTHORED: Init
       #Device.InitCount := #Device.InitCount + 1;
       // ---- GENERATED: reaction end
   END_IF;
   IF #Core.EvCommandStart THEN
       #LatchedParCmd := #ParCmd;
       CASE #Core.Command OF
           1:
               "FRK_Start"(Core := #Core,
                           Status := #Status,
                           Supported := TRUE,
                           Timeout := #ParCfg.Timeout,
                           Label := 'Finish');
           2:
               "FRK_Start"(Core := #Core,
                           Status := #Status,
                           Supported := TRUE,
                           Timeout := #ParCfg.Timeout,
                           Label := 'Wait');
           3:
               "FRK_Start"(Core := #Core,
                           Status := #Status,
                           Supported := TRUE,
                           Timeout := #ParCfg.Timeout,
                           Label := 'Hold');
           4:
               "FRK_Start"(Core := #Core,
                           Status := #Status,
                           Supported := TRUE,
                           Timeout := #ParCfg.Timeout,
                           Label := 'Fault');
           5:
               "FRK_Start"(Core := #Core,
                           Status := #Status,
                           Supported := TRUE,
                           Timeout := #ParCfg.Timeout,
                           Label := 'Pending');
           6:
               "FRK_Start"(Core := #Core,
                           Status := #Status,
                           Supported := TRUE,
                           Timeout := #ParCfg.Timeout,
                           Label := 'Instant');
           7:
               "FRK_Start"(Core := #Core,
                           Status := #Status,
                           Supported := TRUE,
                           Timeout := #ParCfg.Timeout,
                           Label := 'Adopt');
           ELSE
               "FRK_Start"(Core := #Core,
                           Status := #Status,
                           Supported := FALSE,
                           Timeout := T#0ms,
                           Label := '');
       END_CASE;
   END_IF;
   IF #Core.EvCommandStart THEN
       // ---- AUTHORED: CommandStart
       #Device.StartCount := #Device.StartCount + 1;
       #Device.Ordered := #Device.InitCount = 1;
       // ---- GENERATED: reaction end
   END_IF;
   // ---- AUTHORED: cyclic management
   #Device.CyclicCount := #Device.CyclicCount + 1;
   IF #Hal.BackgroundFault THEN
       "FRK_Fault"(Core := #Core,
                   Status := #Status,
                   ReasonCode := 2901,
                   Description := WSTRING#'test.background');
   END_IF;
   // ---- GENERATED: end management
   "FRK_RouteAbort"(Core := #Core,
                    Abort := #Abort);
   IF #Core.EvAbort THEN
       // ---- AUTHORED: Abort
       #Device.AbortCount := #Device.AbortCount + 1;
       // ---- GENERATED: reaction end
   END_IF;
   IF #Core.EvAbortInError THEN
       // ---- AUTHORED: AbortInError
       #Device.ErrorAbortCount := #Device.ErrorAbortCount + 1;
       // ---- GENERATED: reaction end
   END_IF;
   IF #Core.Dispatch AND #Core.RegIndex > 0 AND NOT "FRK_Registry".Fault THEN
       // ---- AUTHORED: dispatch
       #Device.DispatchCount := #Device.DispatchCount + 1;
       #Device.SeenValue := #LatchedParCmd.Value;
       CASE #Core.Command OF
           1:
               IF #Hal.Finish THEN
                   #OutCmd.Result := #LatchedParCmd.Value;
                   "FRK_Complete"(Core := #Core,
                                  Status := #Status);
               END_IF;
           2:
               #Device.SeenValue := #LatchedParCmd.Value;
           3:
               IF NOT #Hal.Permit THEN
                   "FRK_Hold"(Core := #Core,
                              Status := #Status,
                              ReasonCode := 2003,
                              Description := WSTRING#'test.permit');
               ELSIF #Hal.Finish THEN
                   "FRK_Complete"(Core := #Core,
                                  Status := #Status);
               END_IF;
           4:
               "FRK_Fault"(Core := #Core,
                           Status := #Status,
                           ReasonCode := 2901,
                           Description := WSTRING#'test.first');
               "FRK_Fault"(Core := #Core,
                           Status := #Status,
                           ReasonCode := 2001,
                           Description := WSTRING#'test.second');
           5:
               "FRK_Pending"(Core := #Core,
                             Status := #Status,
                             Diag := #Hal.Diag);
               "FRK_Pending"(Core := #Core,
                             Status := #Status,
                             Diag := #Hal.LaterDiag);
           6:
               "FRK_Complete"(Core := #Core,
                              Status := #Status);
           7:
               "FRK_AdoptFault"(Core := #Core,
                                Status := #Status,
                                Diag := #Hal.Diag);
           ELSE
               "FRK_Fault"(Core := #Core,
                           Status := #Status,
                           ReasonCode := 2008,
                           Description := WSTRING#'std.error.unsupportedHmiRequest');
       END_CASE;
       // ---- GENERATED: end dispatch
   END_IF;
   "FRK_End"(Core := #Core,
             Status := #Status,
             Busy => #Busy,
             Done => #Done,
             Error => #Error,
             Aborted => #Aborted,
             Held => #Held,
             ErrorID => #ErrorID,
             Timing => #Timing);
   // ---- AUTHORED: unconditional cyclic/derived data
   #Device.Sample := #Hal.Sample;
   #Device.Output := #Core.Exec = 1 AND NOT #Core.Held AND #Hal.Permit;
   #OutImm := #Device;
   // ---- GENERATED: frame end
END_FUNCTION_BLOCK

FUNCTION_BLOCK "FB_SatelliteUnit"   // FB4, SCL
{ S7_Optimized_Access := 'TRUE' }
VERSION : 0.1
// Generated frame v0.6; change the declaration, then regenerate.
// stored: AutoNumber true, IsIECCheckEnabled false, IsRetainMemResEnabled false, MemoryReserve 100, SetENOAutomatically false, UDAEnableTagReadback false
   VAR_INPUT
      Execute { ExternalWritable := 'False'} : Bool;
      Abort { ExternalWritable := 'False'} : Bool;
      Command { ExternalWritable := 'False'} : DInt;
      ParCfg { ExternalWritable := 'False'} : "ST_DeclarationParCfg";
      ParCmd { ExternalWritable := 'False'} : "ST_DeclarationParCmd";
      ParentIndex { ExternalAccessible := 'False'; ExternalVisible := 'False'; ExternalWritable := 'False'} : DInt;
      Startup { ExternalAccessible := 'False'; ExternalVisible := 'False'; ExternalWritable := 'False'} : Bool;
   END_VAR
   VAR_OUTPUT
      Busy { ExternalWritable := 'False'} : Bool;
      Done { ExternalWritable := 'False'} : Bool;
      Error { ExternalWritable := 'False'} : Bool;
      Aborted { ExternalWritable := 'False'} : Bool;
      Held { ExternalWritable := 'False'} : Bool;
      ErrorID { ExternalWritable := 'False'} : DWord;
      Timing { ExternalWritable := 'False'} : "ST_ModuleTiming";
      OutCmd { ExternalWritable := 'False'} : "ST_DeclarationOutCmd";
      OutImm { ExternalWritable := 'False'} : "ST_UnitProbeImm";
   END_VAR
   VAR_IN_OUT
      Hal : "ST_SatelliteUnitHal";
   END_VAR
   VAR
      Status { ExternalWritable := 'False'; S7_SetPoint := 'True'} : "ST_ModuleStatus";
      Core { ExternalAccessible := 'False'; ExternalVisible := 'False'; ExternalWritable := 'False'; S7_SetPoint := 'True'} : "FRK_Core";
      LatchedParCmd { ExternalAccessible := 'False'; ExternalVisible := 'False'; ExternalWritable := 'False'; S7_SetPoint := 'True'} : "ST_DeclarationParCmd";
      Device { ExternalAccessible := 'False'; ExternalVisible := 'False'; ExternalWritable := 'False'; S7_SetPoint := 'True'} : "ST_UnitProbeDevice";
      Unit { ExternalAccessible := 'False'; ExternalVisible := 'False'; ExternalWritable := 'False'; S7_SetPoint := 'True'} : "FRK_Unit";
      HmiRequest { S7_SetPoint := 'True'} : "ST_HmiRequest";
      ModePolicy { ExternalAccessible := 'False'; ExternalVisible := 'False'; ExternalWritable := 'False'; S7_SetPoint := 'True'} : Array[0..6] of "ST_ModePolicy";
      Access { ExternalWritable := 'False'; S7_SetPoint := 'True'} : "FRK_Access";
      HmiResponse { ExternalWritable := 'False'; S7_SetPoint := 'True'} : "ST_HmiResponse";
      ConfigRev { ExternalWritable := 'False'} : UDInt;
      ConfigCursor { ExternalAccessible := 'False'; ExternalVisible := 'False'; ExternalWritable := 'False'; S7_SetPoint := 'True'} : "FRK_ConfigCursor";
      Part { ExternalWritable := 'False'; S7_SetPoint := 'True'} : "ST_PartContext";
      History { ExternalWritable := 'False'; S7_SetPoint := 'True'} : Array[1..16] of "ST_Diagnostic";
      HistoryHead { ExternalWritable := 'False'} : Int;
      ModeActivePublished { ExternalWritable := 'False'} : DInt;
      RunningPublished { ExternalWritable := 'False'} : Bool;
      StopPendingPublished { ExternalWritable := 'False'} : Bool;
      SupportedModesPublished { ExternalWritable := 'False'} : Array[0..6] of Bool;
      GoodCount { ExternalWritable := 'False'} : UDInt;
      NokCount { ExternalWritable := 'False'} : UDInt;
      ReworkCount { ExternalWritable := 'False'} : UDInt;
      NokReason { ExternalWritable := 'False'} : DInt;
      Cell { ExternalWritable := 'False'; S7_SetPoint := 'True'} : "FB_DeclarationCell";
      Inner { ExternalWritable := 'False'; S7_SetPoint := 'True'} : "FB_InnerUnit";
   END_VAR
   VAR_TEMP
      InstancePath : WString[254];
      RouteMatched : Bool;
      ManualMatched : Bool;
   END_VAR
   VAR CONSTANT
      EXEC_READY : DInt := 0;
      MODULE_TIER : DInt := 1;
   END_VAR
BEGIN

